(* IEC 61131-3 sources: volt/packages/volt-lsp-iec/test-corpus/bakon-nano/Device/Plc Logic/Application/Library Manager/L_TS2P_TechModulesSynchronizingCamming (part 2) *)

(* ---- L_TS2P_CALCULATETARGETPOS.pou ---- *)
FUNCTION_BLOCK L_TS2P_CALCULATETARGETPOS
VAR_INPUT
	XRESET : BOOL;
	XENABLE : BOOL;
	XEXECUTENEXTCUT : BOOL;
	XEXECUTEFIRSTCUT : BOOL;
	XSETCUTTINGLENGTHINSTANT : BOOL;
	XTPNOTVALID : BOOL;
	XEXECUTEGAP : BOOL;
	XRESUMETARGETPOS : BOOL;
	XSTARTFLYINGSAW : BOOL;
	ETMSTATE : L_TB2P_States;
	XSYNCININSTANT : BOOL;
	XSETMATERIALCOUNTER : BOOL;
	LRMATERIALCOUNTER : LREAL;
	LRDELTAMATERIALPOS : LREAL;
	LRSLAVEPOS : LREAL;
	LRCUTTINGLENGTH : LREAL;
	LRMARKSENSORPOS : LREAL;
	LRGAP : LREAL;
	LRMARKPOSITION : LREAL;
	XLOADTOTALCUTTINGLENGTH : BOOL;
	LRLOADTOTALCUTTINGLENGTH : LREAL;
	XLOADTARGETPOS : BOOL;
	LRLOADTARGETPOS : LREAL;
	EMODE : L_TS2P_FlyingSawMode;
	LRVELINMASTER : LREAL;
	LRACCDIST : LREAL;
	LRACCTIME : LREAL;
	LRTASKCYCLETIME : LREAL;
	XEMPTYSTACK : BOOL;
	XSYNCHRONIZED : BOOL;
	XINPOSITION : BOOL;
END_VAR
VAR_OUTPUT
	XEXECUTEGAPOUT : BOOL;
	LRTARGETPOS : LREAL;
	LRTARGETPOS_OUT : LREAL;
	LRTOTALPRODUCTLENGTH : LREAL;
	XCUTTINGLENGTHVALID : BOOL;
	LRACTIVECUTTINGLENGTH : LREAL;
END_VAR
VAR
	LROFFSET_INT : LREAL;
	XGAPREQUESTED : BOOL;
	LRDELTAMATERIALPOS_INT : LREAL;
	LRTOLERANCE : LREAL;
	LROFFSETOUT_INT : LREAL;
	LRGAPTOTAL_INT : LREAL;
	XSYNCININSTANT_LOCK : BOOL;
	XENABLE_OLD : BOOL;
	XSYNCININSTANT_OLD : BOOL;
	LRMATERIALCOUNTER_OLD : LREAL;
	XEXECUTENEXTCUT_OLD : BOOL;
	XEXECUTEGAP_OLD : BOOL;
	XEXECUTEFIRSTCUT_OLD : BOOL;
	EMODE_OLD : WORD;
	ETMSTATE_OLD : L_TB2P_States;
	XTPNOTVALID_OLD : BOOL;
	XSETCUTTINGLENGTHINSTANT_OLD : BOOL;
	XSETMATERIALCOUNTER_OLD : BOOL;
	LRMARKPOSITION_OLD : LREAL;
END_VAR
END_FUNCTION_BLOCK

(* ---- L_TS2P_CALCULATETPCOMPENSATIONFACTOR.pou ---- *)
FUNCTION_BLOCK L_TS2P_CALCULATETPCOMPENSATIONFACTOR
VAR_OUTPUT
	LRFACTOR : LREAL;
	LRCOMPENSATIONCYCLES : LREAL;
END_VAR
VAR_IN_OUT
	TPAXIS : AXIS_REF;
END_VAR
VAR
	LRSETPOSARRAY : ARRAY [0..15] OF LREAL;
	BYCOUNTER : BYTE;
	LRTEMP : LREAL;
	LRPOSDIFF : LREAL;
	LRSETACTDIFF : LREAL;
	XERRORINVALIDAXIS : BOOL;
	LRSETPOS : LREAL;
	LRACTPOS : LREAL;
	LRCYCLELENGTH : LREAL;
	LRADDITIONALCORRECTION : LREAL;
	LRTEMP2 : LREAL;
	XINCREMENTCYCLES : BOOL;
END_VAR
END_FUNCTION_BLOCK

METHOD SEARCHARRAY
END_METHOD

(* ---- L_TS2P_CALCULATETPONMATERIALPOS.pou ---- *)
FUNCTION_BLOCK L_TS2P_CALCULATETPONMATERIALPOS
VAR_INPUT
	XENABLE : BOOL;
	BYTASKCYCLEDELAY : BYTE := 4;
	XMARKRECEIVE : BOOL;
	LRMARKSENSORPOS : LREAL;
	LRACTMARKPOSIN : LREAL;
	LRCYCPOSTPAXIS : LREAL;
	LRCYCVELTPAXIS : LREAL;
	LRCYCLELENGTHTPAXIS : LREAL;
	LRCYCLELENGTHTARGETAXIS : LREAL;
	LRTASKCYCLETIME : LREAL;
	XRESETMARKSTACK : BOOL;
	LRMATERIALCOUNTER : LREAL;
	LRUPPERLIMITWORKINGRANGE : LREAL;
	LRLOWERLIMITWORKINGRANGE : LREAL;
	LRFACTOR : LREAL;
	LRCOMPVELFACTOR : LREAL;
	XSCIPTONEXTPOSOUT : BOOL;
	XSYNCININSTANT : BOOL;
	XEXECUTEFIRSTCUT : BOOL;
END_VAR
VAR_OUTPUT
	LRTPPOSOUT : LREAL;
	XEXECUTEFIRSTCUT_OLD : BOOL;
	LRTPACTTIMESTAMP : LREAL;
	XFULL : BOOL;
	WMARKPOSITIONVALID : WORD;
	WININDEX : WORD;
	ALRMARKPOSITIONARRAY : ARRAY [0..15] OF LREAL := [0, 0, 0, 0, 0, 0, 0, 0, 0, 0, 0, 0, 0, 0, 0, 0];
	ALRTIMESTAMPARRAY : ARRAY [0..15] OF LREAL;
	XEMPTY : BOOL := TRUE;
	WOUTINDEX : WORD;
	BYREMAINMARKSTACK : BYTE := 15;
	XTPRECEIVED : BOOL;
	XMARKRECEIVED : BOOL;
	XTPPOSVALID : BOOL;
	BYCOUNTEROUT : BYTE;
	XERROR : BOOL;
END_VAR
VAR
	R_TRIG1 : R_TRIG;
	LRTIMESTAMP : LREAL;
	BYTPIDLEINDEX : BYTE;
	BYTPACTINDEX : BYTE;
	ALRPOSITION : ARRAY [0..15] OF LREAL;
	BYTPPREVINDEX : BYTE;
	BYTMP : BYTE;
	XSKIPTONEXTPOS : BOOL;
	WTESTCOUNTER : WORD;
	XTEST : BOOL;
	XWAIT : BOOL;
	WCOUNTINVALIDTIMESTAMP : WORD;
	LRDISTINACTMASTER : LREAL;
	BYTEST : BYTE;
	LRMARKPOSITIONDIFF : LREAL;
	LRMARKPOSITIONDIFF2 : LREAL;
	LRPOSFIFOX : ARRAY [1..20] OF LREAL := [10(0)];
	LRPOSFIFOREG : ARRAY [1..20] OF LREAL := [10(0)];
	BYCOUNTER : BYTE := 1;
	LRSTACKDIFFERENCE : LREAL;
	LRTPDELTAINMS : LREAL;
	LRDELTAPCT : LREAL;
	LRTEMP : LREAL;
	IDIRECTION : INT;
	LRACTMARKPOSIN_OLD : LREAL;
	R_TRIG2 : R_TRIG;
	DWSTATE : DWORD;
	WSTOREDPOSVALUES : WORD;
	LRACTMARKPOSIN_INT : LREAL;
	XSYNCININSTANT_OLD : BOOL;
	XWAIT_OLD : BOOL;
	XRESETMARKSTACK_OLD : BOOL;
	BYCNT : BYTE;
	BYSTEPPER : BYTE;
END_VAR
END_FUNCTION_BLOCK

METHOD SEARCHINSTACKNEGATIVE
END_METHOD

METHOD SEARCHINSTACKPOSITIVE
END_METHOD

(* ---- L_TS2P_CAMCREATOR.pou ---- *)
FUNCTION_BLOCK L_TS2P_CAMCREATOR
VAR_INPUT
	XENABLEINTERNALCAMTABLE : BOOL;
	XEXECUTE : BOOL;
	PCAMPOINTS : POINTER TO L_MC2P_CamDataXYVA;
	INUMOFPOINTS : INT;
	LRMASTERMAXVEL : LREAL;
	LRMASTERMAXACC : LREAL;
	LRMASTERSCALING : LREAL := 1;
	LRSLAVESCALING : LREAL := 1;
END_VAR
VAR_OUTPUT
	XINTERNALCAMTABLELACTIVE : BOOL;
	XERROR : BOOL;
	EERRORID : L_IE1P_Error;
	XBUSY : BOOL;
	XDONE : BOOL;
	CAMTABLEOUT : MC_CAM_REF;
	LRSLAVEMAXPOS : LREAL;
	LRSLAVEMINPOS : LREAL;
	LRSLAVEMAXVEL : LREAL;
	LRSLAVEMINVEL : LREAL;
	LRSLAVEMAXACC : LREAL;
	LRSLAVEMINACC : LREAL;
END_VAR
VAR_IN_OUT
	SLAVE : AXIS_REF;
END_VAR
VAR
	EFMSTATE : L_MB1P_States := L_MB1P_States.INIT;
	SMC_CAMBOUNDS1 : L_MC2P_BoundsCam;
	SMC_CAMBOUNDSINIT : L_MC2P_BoundsCam;
	CAMREF : L_MC2P_CamRefFromStruct;
	PCAMPOINTS_INT : POINTER TO L_MC2P_CamDataXYVA;
	INUMOFPOINTS_INT : INT;
	XINTERNALCONTROL : BOOL;
	XEXECUTE_OLD : BOOL;
	ASCCAMPOINTS : ARRAY [0..30] OF L_MC2P_CamDataXYVA;
	XINVALIDCAMTABLE : BOOL;
	XVISUACTIVE : BOOL := TRUE;
	DIFRAME : DINT;
	DIFRAME_OLD : DINT;
	ARVISPOINTLINES : ARRAY [1..10] OF L_MC2P_CamDataXYVA;
	IVISUTABLESETPOS : INT := 0;
	IVISUTABLESETPOS_OLD : INT := 0;
	IVISUTABLEMAXPOS : INT := 30;
	IVISSHOWLINESNO : INT;
	XVISPOINTMIN : BOOL;
	XVISPOINTMAX : BOOL;
	XVISUSETPOSUP : BOOL;
	XVISUSETPOSDOWN : BOOL;
	XVISUSETPOSUP_OLD : BOOL;
	XVISUSETPOSDOWN_OLD : BOOL;
	XSCROLBUTTENACTIVE : BOOL;
	TSETTIME : TIME := TIME#400ms;
	TON_SCROLBUTTEN : TON;
END_VAR
END_FUNCTION_BLOCK

METHOD CALL_CAMBOUNDS
VAR_IN_OUT
	SLAVE : AXIS_REF;
END_VAR
END_METHOD

METHOD CALL_CAMREF
END_METHOD

METHOD CALL_CAMTABLEEQUIDISTANT
END_METHOD

METHOD CALL_CAMTABLENONEQUIDISTANT
END_METHOD

METHOD CALL_CAMTABLEPOLYNOMIAL
END_METHOD

METHOD CALL_ERRORHANDLER
END_METHOD

METHOD CALL_FBMETHODS
VAR_IN_OUT
	SLAVE : AXIS_REF;
END_VAR
END_METHOD

METHOD CALL_INTERNALCTRL
END_METHOD

METHOD CALL_OUTPUT
END_METHOD

METHOD CALL_RESETCOMMANDS
VAR_IN_OUT
	SLAVE : AXIS_REF;
END_VAR
END_METHOD

METHOD CALL_RESETOUTPUT
END_METHOD

METHOD CALL_STATEMACHINE
END_METHOD

METHOD CALL_VIS_TON_SCROLBUTTEN
END_METHOD

METHOD CALL_VISUTABCTRL
END_METHOD

METHOD CALL_VISUUPDATETAB
END_METHOD

METHOD DISABALE_VISU
END_METHOD

METHOD ENABLE_VISU
END_METHOD

METHOD CALL_S000_CYCLIC
END_METHOD

METHOD CALL_S001_INIT
END_METHOD

METHOD CALL_S002_READY
END_METHOD

(* ---- L_TS2P_CAMTABLEINFO.pou ---- *)
FUNCTION_BLOCK L_TS2P_CAMTABLEINFO
VAR_INPUT
	XENABLE : BOOL;
	CAMTABLE : MC_CAM_REF;
	LRMASTERMAXVEL : LREAL := 100;
	LRMASTERMAXACC : LREAL := 1000;
	LRMASTERSCALING : LREAL := 1;
	LRSLAVESCALING : LREAL := 1;
END_VAR
VAR_OUTPUT
	XBUSY : BOOL;
	XDONE : BOOL;
	XCAMTABLEVALID : BOOL;
	LRMASTERSTARTPOS : LREAL;
	LRMASTERENDPOS : LREAL;
	LRSLAVESTARTPOS : LREAL;
	LRSLAVEENDPOS : LREAL;
	LRSLAVEMAXPOS : LREAL;
	LRSLAVEMINPOS : LREAL;
	LRSLAVEMAXVEL : LREAL;
	LRSLAVEMINVEL : LREAL;
	LRSLAVEMAXACC : LREAL;
	LRSLAVEMINACC : LREAL;
END_VAR
VAR_IN_OUT
	SLAVEAXIS : AXIS_REF;
END_VAR
VAR
	ESTATE : L_MB1P_States := L_MB1P_States.INIT;
	CAMTABLE_INT : MC_CAM_REF;
	PCAMDATA_INT : POINTER TO L_MC2P_CamData;
	LRMASTERMAXVEL_INT : LREAL := 0;
	LRMASTERMAXACC_INT : LREAL := 0;
	LRMASTERSCALING_INT : LREAL := 0;
	LRSLAVESCALING_INT : LREAL := 0;
	XENABLE_OLD : BOOL;
	SMC_CAMBOUNDS1 : L_MC2P_BoundsCam;
	XCALCNEWVALUES : BOOL;
END_VAR
END_FUNCTION_BLOCK

METHOD CALC_STARTENDVALUES
END_METHOD

METHOD CALL_CAMBOUNDS
END_METHOD

METHOD CALL_FBMETHODS
END_METHOD

METHOD CALL_OUTPUT
END_METHOD

METHOD CALL_RESETCOMMANDS
END_METHOD

METHOD CALL_RESETOUTPUT
END_METHOD

METHOD CALL_STATEMACHINE
END_METHOD

METHOD GET_XCALCNEWVALUES : BOOL
END_METHOD

METHOD GET_XCRITICALCYCLE : BOOL
END_METHOD

(* ---- L_TS2P_CONDITIONLIMITERSYNCIN.pou ---- *)
FUNCTION_BLOCK L_TS2P_CONDITIONLIMITERSYNCIN EXTENDS L_UBUP_ConditionBase
VAR_INPUT
	ESYNCDIRECTION : L_TS2P_SyncDirection;
	DWLIMITERCONTROL : DWORD;
END_VAR
VAR_OUTPUT
	XDIRECTIONDISABLED : BOOL;
	XINVALIDINPUT : BOOL;
END_VAR
VAR_IN_OUT
	AXIS : AXIS_REF;
END_VAR
END_FUNCTION_BLOCK

METHOD VERIFY : BOOL
VAR_OUTPUT
	XCONDITIONERROR : BOOL;
	EERRORIDPROPOSED : L_IE1P.L_IE1P_Error;
END_VAR
END_METHOD

(* ---- L_TS2P_CONDITIONLOCKTOCAM.pou ---- *)
FUNCTION_BLOCK L_TS2P_CONDITIONLOCKTOCAM EXTENDS L_UBUP_ConditionBase
VAR_IN_OUT
	SCPAR : L_TS2P_scPar_TM_FlexCam;
END_VAR
END_FUNCTION_BLOCK

METHOD VERIFY : BOOL
VAR_OUTPUT
	XCONDITIONERROR : BOOL;
	EERRORIDPROPOSED : L_IE1P.L_IE1P_Error;
END_VAR
END_METHOD

(* ---- L_TS2P_CONDITIONSYNCPARAMETER.pou ---- *)
FUNCTION_BLOCK L_TS2P_CONDITIONSYNCPARAMETER EXTENDS L_UBUP_ConditionBase
VAR_IN_OUT
	SCPAR : L_TS2P_scPar_TM_SyncPosBase;
END_VAR
END_FUNCTION_BLOCK

METHOD VERIFY : BOOL
VAR_OUTPUT
	XCONDITIONERROR : BOOL;
	EERRORIDPROPOSED : L_IE1P.L_IE1P_Error;
END_VAR
END_METHOD

(* ---- L_TS2P_CONDITIONVALIDCAMTABLE.pou ---- *)
FUNCTION_BLOCK L_TS2P_CONDITIONVALIDCAMTABLE EXTENDS L_UBUP_ConditionBase
VAR_INPUT
	WSETCAMTABLE : WORD;
	CAMTABLE1 : MC_CAM_REF;
	CAMTABLE2 : MC_CAM_REF;
	CAMTABLE3 : MC_CAM_REF;
	CAMTABLE4 : MC_CAM_REF;
END_VAR
END_FUNCTION_BLOCK

METHOD VERIFY : BOOL
VAR_OUTPUT
	XCONDITIONERROR : BOOL;
	EERRORIDPROPOSED : L_IE1P.L_IE1P_Error;
END_VAR
END_METHOD

(* ---- L_TS2P_CROSSCUTTERSTATE.pou ---- *)
FUNCTION_BLOCK L_TS2P_CROSSCUTTERSTATE EXTENDS L_TB2P_TechModuleBase
VAR_INPUT
	XENABLE : BOOL;
	XENABLEOPERATION : BOOL;
	XRESETERROR : BOOL;
	XQSPAPPLICATION : BOOL;
	XABORT : BOOL;
	XJOGPOS : BOOL;
	XJOGNEG : BOOL;
	XHOMEEXECUTE : BOOL;
	LROVERRIDE : LREAL := 1;
	SCCTRLBASICMOTION : L_TB2P_scCtrlBasicMotion;
	SCPAR : L_TS2P_scPar_CrossCutterState;
	SCACCESSPOINTS : L_TS2P_scAP_CrossCutterState;
	MASTERVALUES : L_MC1P_IAXIS_REF_MASTERVALUES;
	XEXECUTEMOVETOPARKPOS : BOOL;
	XSYNCIN : BOOL;
	XHOLDINPARKPOS : BOOL;
	LRPRODUCTLENGTH : LREAL;
	LROVERSPEED : LREAL;
	LRSETOFFSETPOSX : LREAL;
	XTRIMPOS : BOOL;
	XTRIMNEG : BOOL;
	XTRIMRESET : BOOL;
	SCTPRECDATA_MARKSENSOR : L_MC1P_TpReceiveData;
	SCTPRECDATA_TOOLSENSOR : L_MC1P_TpReceiveData;
	XTEACHMARKWINDOW : BOOL;
	XTEACHMARKWINDOWTOOL : BOOL;
	XGEARFACTORCORR : BOOL;
	XGEARFACTORCORRHOLD : BOOL;
END_VAR
VAR_OUTPUT
	XREADYFOROPERATION : BOOL;
	XOPERATIONENABLED : BOOL;
	XREADYFORMOTION : BOOL;
	XERROR : BOOL;
	XWARNING : BOOL;
	EERRORID : L_IE1P_Error;
	XSTOACTIVE : BOOL;
	XQSPACTIVE : BOOL;
	XABORTBUSY : BOOL;
	XABORTDONE : BOOL;
	XJOGGINGBUSY : BOOL;
	XHOMINGBUSY : BOOL;
	XHOMINGDONE : BOOL;
	XISHOMED : BOOL;
	ETMSTATE : L_TB2P_States;
	SCSTATUSBASICMOTION : L_TB2P_scStatusBasicMotion;
	LRACTVEL : LREAL;
	LRSETVELOUT : LREAL;
	LRACTPOS : LREAL;
	LRSETPOSOUT : LREAL;
	LRACTFOLLOWINGERROR : LREAL;
	SCSIGNALFLOW : L_TS2P_scSF_CrossCutterState;
	XSYNCHRONISED : BOOL;
	XACCDECSYNC : BOOL;
	XOFFSETTRIMACTIVE : BOOL;
	XINPARKPOS : BOOL;
	XHOLDINPARKPOSACTIVE : BOOL;
	XCUTDONE : BOOL;
	XCUTTINGACTIVE : BOOL;
	LRACTCUTLENGTH : LREAL;
	LROFFSETTOTAL : LREAL;
	XTRQCTRLACTIVE : BOOL;
	LRSETMARKCORROUT : LREAL;
	XMARKWINDOWTEACHED : BOOL;
	LRGEARFACTORCORR : LREAL;
	LRSETTOOLCORROUT : LREAL;
	XMARKWINDOWTEACHEDTOOL : BOOL;
END_VAR
VAR_IN_OUT
	AXIS : AXIS_REF;
END_VAR
VAR
	TM_INT : L_TS2P_TM_CrossCutterState := STRUCT(ModuleHandler := ModuleHandler);
	SCPAR_INT : L_TS2P_scPar_CrossCutterState;
	_UICALLMFUNIDXINPUT : UINT := 1;
	_UICALLMFUNIDXOUTPUT : UINT := 1;
	_MCCALL : L_UM1P_MCCall;
	_ASCINPUT : ARRAY [1.._MCCall.c_BufferDepthInput] OF L_TS2P_CrossCutterStateIn;
	_ASCOUTPUT : ARRAY [1.._MCCall.c_BufferDepthOutput] OF L_TS2P_CrossCutterStateOut;
	_ASCPARCORE : ARRAY [1.._MCCall.c_BufferDepthInput] OF L_TS2P_scPar_CrossCutterState;
	_ASCACCESSPOINTSCORE : ARRAY [1.._MCCall.c_BufferDepthInput] OF L_TS2P_scAP_CrossCutterState;
	_ASCSIGNALFLOWCORE : ARRAY [1.._MCCall.c_BufferDepthOutput] OF L_TS2P_scSF_CrossCutterState;
	_SCINPUTVISU : L_TS2P_CrossCutterStateIn;
	_PSCINPUTVISU : POINTER TO L_TS2P_CrossCutterStateIn := ADR(_scInputVisu);
	_PSCOUTPUTVISU : POINTER TO L_TS2P_CrossCutterStateOut := ADR(_ascOutput[1]);
	_PSCPARVISU : POINTER TO L_TS2P_scPar_CrossCutterState := ADR(scPar_int);
	ITFITECHMODULEINTERNAL : L_TB2P_ITechModuleInternal;
	LRJERKDEC : LREAL;
	LRJOGGINGJERKDEC : LREAL;
	REMAININGTIMEOFPROFILE : LREAL;
	REMAININGTIMEOFPROFILEAVAILABLE : BOOL;
END_VAR
END_FUNCTION_BLOCK

METHOD GET_PAP : POINTER TO L_TB2P_scAP_TM_MotionControl
END_METHOD

METHOD GET_PPAR : POINTER TO L_TB2P_scPar_TM_MotionControl
END_METHOD

METHOD GET_PSF : POINTER TO L_TB2P_scSF_TM_MotionControl
END_METHOD

METHOD CALLFUNCTION
VAR_INPUT
	UIINPUTDATAIDX : UINT;
	UIOUTPUTDATAIDX : UINT;
END_VAR
END_METHOD

METHOD COPYINPUTS : BOOL
VAR_INPUT
	IDX : WORD;
END_VAR
END_METHOD

METHOD COPYOUTPUTS : BOOL
VAR_INPUT
	IDX : WORD;
END_VAR
END_METHOD

METHOD FUNCTIONWASCALLEDTWICE : BOOL
VAR_INPUT
	IDX : WORD;
END_VAR
END_METHOD

METHOD HANDLESTANDARDCALL : BOOL
END_METHOD

METHOD SYNCOUTPUTS
VAR_INPUT
	UICOPYOUTPUTFROMIDX : UINT;
	UICOPYOUTPUTTOIDX : UINT;
END_VAR
END_METHOD

METHOD CALL_INTERNALCTRL
END_METHOD

(* ---- L_TS2P_DISTCORRECTIONWINDOW.pou ---- *)
FUNCTION_BLOCK L_TS2P_DISTCORRECTIONWINDOW
VAR_INPUT
	XENABLE : BOOL;
	XENABLEPOSITION : BOOL;
	LRCYCSETPOSMASTER : LREAL;
	LRCYCLELENGTHMASTER : LREAL;
	LRCYCSETVEL : LREAL;
	XLOADSTARTPOS : BOOL;
	LRSTARTPOS : LREAL;
	XTPRECEIVEDIN : BOOL;
	LRSETCORRECTION : LREAL;
	XCORRWINDOWINXUNITS : BOOL;
	LRSETUPPERWINDOW : LREAL;
	LRSETLOWERWINDOW : LREAL;
	LRCYCPOSFEEDBACK : LREAL;
	DNSETNUMERATORAXISY : DWORD := 1;
	DNSETDENOMINATORAXISY : DWORD := 1;
	LRSETCYCLELENGTHX : LREAL;
	LRSETCYCLELENGTHY : LREAL;
END_VAR
VAR_OUTPUT
	XBUSY : BOOL;
	XCORRECTIONBUSY : BOOL;
	LRSETPOSOUT : LREAL;
	LRSETINTEGRATEDPOSITION : LREAL;
	LRSETPOSCORROUT : LREAL;
	LRSETPOSCORRRESIDUALOUT : LREAL;
	LRDELTAPOSCORROUT : LREAL;
	XCORRNEXTCYCLE : BOOL;
	XERROR : BOOL;
	EERRORID : L_IE1P_Error;
END_VAR
VAR
	LRDELTAPOSTOTAL : LREAL;
	LRMASTERDISTANCE : LREAL;
	LRPOSITIONSET : LREAL;
	LRPOSITIONNORMED : LREAL;
	LRPOSITIONOUTNORMED : LREAL;
	LRDELTAPOSCORRECTION : LREAL;
	LRPOSITIONSETOLD : LREAL;
	LRPOSITIONSETAXISOUT : LREAL;
	BYSTEPPER : BYTE;
	LRCORRECTIONDISTANCELOCAL : LREAL;
	LRCORRECTIONLOCAL : LREAL;
	L_DIFFERENTIATE : L_MC2P_Differentiate;
	INTEGRATOR : L_MC1P_IntegrateAxis;
	LRDELTAPOSOUT : LREAL;
	XEXECUTECORRECTIONINTERN : BOOL;
	XPOSITIVEDIRECTION : BOOL := FALSE;
	LRCORRECTIONDISTANCE : LREAL;
	LRUPPERWINDOWINTERNAL : LREAL;
	LRLOWERWINDOWINTERNAL : LREAL;
	LRTASKCYCLE : LREAL;
	XCORRECTIONACTIVE : BOOL;
	LRCORRECTIONLOCAL1 : LREAL;
	XTPRECEIVEDOLD : BOOL;
	LRINTEGRATORSPEED : LREAL;
	XWINDOWINCYCLE : BOOL;
	LRDELTAWINDOW : LREAL;
	LRCYCPOSINTOOLINTERNAL : LREAL;
	LRUPPERWINDOWINTERNALDELTA : LREAL;
	LRLOWERWINDOWINTERNALDELTA : LREAL;
	XINIT : BOOL := TRUE;
	XINITOUTOFCORRWINDOW : BOOL := TRUE;
	LRLOWERWINDOWINTERNALOLD : LREAL;
	LRUPPERWINDOWINTERNALOLD : LREAL;
	LRCYCPOSFEEDBACKINT : LREAL;
	XCORRECTIONBUSYOLD : BOOL;
	LRSETPOSCORROUTOLD : LREAL;
	LRCYCPOSINTOOLINTERNAL_CASE : LREAL;
	XWINDOWCHANGEDFLAG : BOOL := FALSE;
	LRCYCLELENGTH_INT : LREAL;
	LROFFSET_INT : LREAL;
	LRCYCPOSINTOOLINTERNAL_0LD : LREAL;
	LRPOSITIONNORMED_OLD : LREAL;
	LRPOSITIONNORMED_DIF : LREAL;
	XPOSCORR : BOOL;
	XTPSTORED_INT : BOOL;
	LRSETCORRECTIONSTORED_INT : LREAL;
	XINCORRWINDOW : BOOL;
	XINCORRWINDOWOLD : BOOL;
	LRSETPOSOUTCOMP : LREAL;
	LRCYCPOSINTOOLINTERNALOLD : LREAL;
	LRDELTAPOSOUTINTERNAL : LREAL;
	BYSTEPPEROLD : BYTE := 0;
	LRCYCSETPOSOLD : LREAL;
	LRCORRECTIONINYUNITS : LREAL;
	LRCORRECTIONDISTANCETEMP : LREAL;
END_VAR
END_FUNCTION_BLOCK

METHOD CALL_INIT
END_METHOD

(* ---- L_TS2P_ELECTRONICGEARBOXBASE.pou ---- *)
FUNCTION_BLOCK L_TS2P_ELECTRONICGEARBOXBASE EXTENDS L_TB2P_TechModuleBase
VAR_INPUT
	XENABLE : BOOL;
	XENABLEOPERATION : BOOL;
	XRESETERROR : BOOL;
	XQSPAPPLICATION : BOOL;
	XABORT : BOOL;
	XJOGPOS : BOOL;
	XJOGNEG : BOOL;
	XHOMEEXECUTE : BOOL;
	LROVERRIDE : LREAL := 1;
	SCCTRLBASICMOTION : L_TB2P_scCtrlBasicMotion;
	SCPAR : L_TS2P_scPar_ElectronicGearboxBase;
	SCACCESSPOINTS : L_TS2P_scAP_ElectronicGearboxBase;
	MASTERVALUES : L_MC1P_IAXIS_REF_MASTERVALUES;
	XSYNCIN : BOOL;
	LRSETBASEVEL : LREAL;
	LRSETOFFSETPOS : LREAL;
	LRSETOFFSETVEL : LREAL;
	XTRIMPOS : BOOL;
	XTRIMNEG : BOOL;
	XTRIMRESET : BOOL;
	XINVERTGEARFACTOR : BOOL;
END_VAR
VAR_OUTPUT
	XREADYFOROPERATION : BOOL;
	XOPERATIONENABLED : BOOL;
	XREADYFORMOTION : BOOL;
	XERROR : BOOL;
	XWARNING : BOOL;
	EERRORID : L_IE1P_Error;
	XSTOACTIVE : BOOL;
	XQSPACTIVE : BOOL;
	XABORTBUSY : BOOL;
	XABORTDONE : BOOL;
	XJOGGINGBUSY : BOOL;
	XHOMINGBUSY : BOOL;
	XHOMINGDONE : BOOL;
	XISHOMED : BOOL;
	ETMSTATE : L_TB2P_States := L_TB2P_States.DISABLED;
	SCSTATUSBASICMOTION : L_TB2P_scStatusBasicMotion;
	LRACTVEL : LREAL;
	LRSETVELOUT : LREAL;
	LRACTPOS : LREAL;
	LRSETPOSOUT : LREAL;
	LRACTFOLLOWINGERROR : LREAL;
	SCSIGNALFLOW : L_TS2P_scSF_ElectronicGearboxBase;
	XSYNCHRONISED : BOOL;
	XACCDECSYNC : BOOL;
	XOFFSETTRIMACTIVE : BOOL;
	XBASEVELOCITYACTIVE : BOOL;
	LROFFSETTOTALVEL : LREAL;
END_VAR
VAR_IN_OUT
	AXIS : AXIS_REF;
END_VAR
VAR
	TM_INT : L_TS2P_TM_ElectronicGearboxBase := STRUCT(ModuleHandler := ModuleHandler);
	SCPAR_INT : L_TS2P_scPar_ElectronicGearboxBase;
	_UICALLMFUNIDXINPUT : UINT := 1;
	_UICALLMFUNIDXOUTPUT : UINT := 1;
	_MCCALL : L_UM1P_MCCall;
	_ASCINPUT : ARRAY [1.._MCCall.c_BufferDepthInput] OF L_TS2P_ElectronicGearboxBaseIn;
	_ASCOUTPUT : ARRAY [1.._MCCall.c_BufferDepthOutput] OF L_TS2P_ElectronicGearboxBaseOut;
	_ASCPARCORE : ARRAY [1.._MCCall.c_BufferDepthInput] OF L_TS2P_scPar_ElectronicGearboxBase;
	_ASCACCESSPOINTSCORE : ARRAY [1.._MCCall.c_BufferDepthInput] OF L_TS2P_scAP_ElectronicGearboxBase;
	_ASCSIGNALFLOWCORE : ARRAY [1.._MCCall.c_BufferDepthOutput] OF L_TS2P_scSF_ElectronicGearboxBase;
	_SCINPUTVISU : L_TS2P_ElectronicGearboxBaseIn;
	_PSCINPUTVISU : POINTER TO L_TS2P_ElectronicGearboxBaseIn := ADR(_scInputVisu);
	_PSCOUTPUTVISU : POINTER TO L_TS2P_ElectronicGearboxBaseOut := ADR(_ascOutput[1]);
	_PSCPARVISU : POINTER TO L_TS2P_scPar_ElectronicGearboxBase := ADR(scPar_int);
	ITFITECHMODULEINTERNAL : L_TB2P_ITechModuleInternal;
	LRJERKDEC : LREAL;
	LRJOGGINGJERKDEC : LREAL;
	REMAININGTIMEOFPROFILE : LREAL;
	REMAININGTIMEOFPROFILEAVAILABLE : BOOL;
END_VAR
END_FUNCTION_BLOCK

METHOD GET_PAP : POINTER TO L_TB2P_scAP_TM_MotionControl
END_METHOD

METHOD GET_PPAR : POINTER TO L_TB2P_scPar_TM_MotionControl
END_METHOD

METHOD GET_PSF : POINTER TO L_TB2P_scSF_TM_MotionControl
END_METHOD

METHOD CALLFUNCTION
VAR_INPUT
	UIINPUTDATAIDX : UINT;
	UIOUTPUTDATAIDX : UINT;
END_VAR
END_METHOD

METHOD COPYINPUTS : BOOL
VAR_INPUT
	IDX : WORD;
END_VAR
END_METHOD

METHOD COPYOUTPUTS : BOOL
VAR_INPUT
	IDX : WORD;
END_VAR
END_METHOD

METHOD FUNCTIONWASCALLEDTWICE : BOOL
VAR_INPUT
	IDX : WORD;
END_VAR
END_METHOD

METHOD HANDLESTANDARDCALL : BOOL
END_METHOD

METHOD SYNCOUTPUTS
VAR_INPUT
	UICOPYOUTPUTFROMIDX : UINT;
	UICOPYOUTPUTTOIDX : UINT;
END_VAR
END_METHOD

METHOD CALL_INTERNALCTRL
END_METHOD

(* ---- L_TS2P_FLEXCAMHIGH.pou ---- *)
FUNCTION_BLOCK L_TS2P_FLEXCAMHIGH EXTENDS L_TB2P_TechModuleBase
VAR_INPUT
	XUSEORIGINAL : BOOL;
	XENABLE : BOOL;
	XENABLEOPERATION : BOOL;
	XRESETERROR : BOOL;
	XQSPAPPLICATION : BOOL;
	XABORT : BOOL;
	XJOGPOS : BOOL;
	XJOGNEG : BOOL;
	XHOMEEXECUTE : BOOL;
	LROVERRIDE : LREAL := 1;
	SCCTRLBASICMOTION : L_TB2P_scCtrlBasicMotion;
	SCPAR : L_TS2P_scPar_FlexCamHigh;
	SCACCESSPOINTS : L_TS2P_scAP_FlexCamHigh;
	MASTERVALUES : L_MC1P_IAXIS_REF_MASTERVALUES;
	XCLUTCHCLOSE : BOOL;
	XLOADCLUTCHPOS : BOOL;
	LRLOADCLUTCHPOS : LREAL;
	XFINDCLUTCHXPOS : BOOL;
	XSYNCIN : BOOL;
	XSYNCPOSRESTORE : BOOL;
	XCAMCHANGEINSTANT : BOOL;
	LRSETOFFSETPOSX : LREAL;
	LRSETOFFSETPOSY : LREAL;
	LRSETSCALINGX : LREAL := 1;
	LRSETSCALINGY : LREAL := 1;
	CAMTABLE1 : MC_CAM_REF;
	CAMTABLE2 : MC_CAM_REF;
	CAMTABLE3 : MC_CAM_REF;
	CAMTABLE4 : MC_CAM_REF;
	WSETCAMTABLE : WORD := 1;
	XCAMSEQUENCER : BOOL;
END_VAR
VAR_OUTPUT
	XREADYFOROPERATION : BOOL;
	XOPERATIONENABLED : BOOL;
	XREADYFORMOTION : BOOL;
	XERROR : BOOL;
	XWARNING : BOOL;
	EERRORID : L_IE1P_Error;
	XSTOACTIVE : BOOL;
	XQSPACTIVE : BOOL;
	XABORTBUSY : BOOL;
	XABORTDONE : BOOL;
	XJOGGINGBUSY : BOOL;
	XHOMINGBUSY : BOOL;
	XHOMINGDONE : BOOL;
	XISHOMED : BOOL;
	ETMSTATE : L_TB2P_States;
	SCSTATUSBASICMOTION : L_TB2P_scStatusBasicMotion;
	LRACTVEL : LREAL;
	LRSETVELOUT : LREAL;
	LRACTPOS : LREAL;
	LRSETPOSOUT : LREAL;
	LRACTFOLLOWINGERROR : LREAL;
	SCSIGNALFLOW : L_TS2P_scSF_FlexCamHigh;
	XCLUTCHACTIVE : BOOL;
	XCLUTCHCLOSED : BOOL;
	XACCDECSYNC : BOOL;
	XSYNCHRONISED : BOOL;
	XMOVETOPARKPOSACTIVE : BOOL;
	XINPARKPOS : BOOL;
	XENDOFPROFILE : BOOL;
	LROFFSETPOSX : LREAL;
	LROFFSETPOSY : LREAL;
	LROFFSETSYNCPOS : LREAL;
	WACTIVECAMTABLE : WORD;
	XCAMSEQUENCERACTIVE : BOOL;
END_VAR
VAR_IN_OUT
	AXIS : AXIS_REF;
END_VAR
VAR
	XINTERNALCONTROLACTIVE_OLD : BOOL;
	ITFCONNECTORFLEXCAM : L_TS2P_IConnectorFlexCam;
	TM_INT : L_TS2P_TM_FlexCam;
	SCPAR_INT : L_TS2P_scPar_FlexCamHigh;
	SCDATA_INT : L_TS2P_scData_TM_FlexCam;
	SCDATASP_INT : L_TS2P_scData_TM_FlexCam;
	XUSEORIGINAL_OLD : BOOL;
	_UICALLMFUNIDXINPUT : UINT := 1;
	_UICALLMFUNIDXOUTPUT : UINT := 1;
	_MCCALL : L_UM1P_MCCall;
	_ASCINPUT : ARRAY [1.._MCCall.c_BufferDepthInput] OF L_TS2P_FlexCamHighIn;
	_ASCOUTPUT : ARRAY [1.._MCCall.c_BufferDepthOutput] OF L_TS2P_FlexCamHighOut;
	_ASCPARCORE : ARRAY [1.._MCCall.c_BufferDepthInput] OF L_TS2P_scPar_FlexCamHigh;
	_ASCACCESSPOINTSCORE : ARRAY [1.._MCCall.c_BufferDepthInput] OF L_TS2P_scAP_FlexCamHigh;
	_ASCSIGNALFLOWCORE : ARRAY [1.._MCCall.c_BufferDepthOutput] OF L_TS2P_scSF_FlexCamHigh;
	_SCINPUTVISU : L_TS2P_FlexCamHighIn;
	_PSCINPUTVISU : POINTER TO L_TS2P_FlexCamHighIn := ADR(_scInputVisu);
	_PSCOUTPUTVISU : POINTER TO L_TS2P_FlexCamHighOut := ADR(_ascOutput[1]);
	_PSCDATAVISU : POINTER TO L_TS2P_scData_TM_FlexCam := ADR(scData_int);
	_PSCPARVISU : POINTER TO L_TS2P_scPar_FlexCamHigh := ADR(scPar_int);
	_PSCAPVISU : POINTER TO L_TS2P_scAP_FlexCamHigh;
	_PSCSFVISU : POINTER TO L_TS2P_scSF_FlexCamHigh;
	ITFBASICMOTIONBASE : L_TB2P.L_TB2P_IBasicMotionBase;
	ITFFLEXCAMEXTENSION : L_TS2P_IFlexCam;
	ITFITECHMODULEINTERNAL : L_TB2P_ITechModuleInternal;
	LRJERKDEC : LREAL;
	LRJOGGINGJERKDEC : LREAL;
	REMAININGTIMEOFPROFILE : LREAL;
	REMAININGTIMEOFPROFILEAVAILABLE : BOOL;
END_VAR
END_FUNCTION_BLOCK

METHOD CALL_ABC
VAR_INPUT
	ITFTECHMODULE : L_TB2P.L_TB2P_IBasicMotionBase;
	XQSPAPPLICATION : BOOL;
	XHALT : BOOL;
	XABORT : BOOL;
	XHOMEEXECUTE : BOOL;
	XJOGPOS : BOOL;
	XJOGNEG : BOOL;
	XFINISHPOSITIONING : BOOL;
	XMOVEVELEXECUTE : BOOL;
	XMOVEABSEXECUTE : BOOL;
	XMOVERELEXECUTE : BOOL;
	XENABLEOPERATION : BOOL;
	XRESETERROR : BOOL;
	XENABLEPOSITIVE : BOOL;
	XENABLENEGATIVE : BOOL;
	XDISABLESWLIMIT : BOOL;
	LROVERRIDE : LREAL;
	LROVERRIDEACC : LREAL;
	LROVERRIDEJERK : LREAL;
	XRESETHOMEPOSITION : BOOL;
	XCONTINUOUSUPDATE : BOOL;
	LRPOS_DIST : LREAL;
	LRVEL : LREAL;
	LRACC : LREAL;
	LRDEC : LREAL;
	LRJERK : LREAL;
	EDIRECTION : L_TB2P.MC_DIRECTION;
	SCHOMEEXTTP : L_TB2P.MC_TRIGGER_REF;
	XHOMEABSSWITCH : BOOL;
	XSPECIALABORTBEHAVIOR : BOOL;
	LRABORTDEC : LREAL;
	LRABORTJERK : LREAL;
END_VAR
VAR_OUTPUT
	XERROR : BOOL;
	EERRORID : L_TB2P.L_IE1P_Error;
	XFUNBUSY : BOOL;
	XFUNDONE : BOOL;
	XFUNCOMMANDABORTED : BOOL;
	EFUNSTATEACT : L_TB2P.L_MC1P_ABC_State;
	ECONTROLMODE : L_TB2P.L_MC1P_ControlMode;
	XISHOMED : BOOL;
	XHWLIMITSWITCHNEG : BOOL;
	XHWLIMITSWITCHPOS : BOOL;
	XSWLIMITENABLED : BOOL;
	XSWLIMITSWITCHNEG : BOOL;
	XSWLIMITSWITCHPOS : BOOL;
	EAXISTYPE : L_TB2P.L_MC1P_DriveType;
	EAXISSTATE : L_TB2P.L_MC1P_AXIS_STATE;
	XSTOACTIVE : BOOL;
	XREADYFOROPERATION : BOOL;
	XOPERATIONENABLED : BOOL;
	XREADYFORMOTION : BOOL;
	XAXISWARNING : BOOL;
	XAXISERROR : BOOL;
	EAXISERRORID : L_TB2P.L_IE1P_Error;
	XDRIVEWARNING : BOOL;
	XDRIVEERROR : BOOL;
	DWDRIVEERRORID : DWORD;
	LRACTPOS : LREAL;
	LRACTVEL : LREAL;
	LRSETPOSOUT : LREAL;
	LRSETVELOUT : LREAL;
	LRACTFOLLOWINGERROR : LREAL;
	XINPOSITION : BOOL;
	XSTANDSTILLSETVELOCITY : BOOL;
	XSTANDSTILLACTVELOCITY : BOOL;
	XCONSTANTVELOCITY : BOOL;
	XACCELERATING : BOOL;
	XDECELERATING : BOOL;
	XDIRECTIONPOSITIVE : BOOL;
	XDIRECTIONNEGATIVE : BOOL;
	XAXISAVAILABLE : BOOL;
END_VAR
VAR_IN_OUT
	AXIS : AXIS_REF;
END_VAR
END_METHOD

METHOD GET_PAP : POINTER TO L_TB2P_scAP_TM_MotionControl
END_METHOD

METHOD GET_PDATA : POINTER TO L_TS2P_scData_TM_FlexCam
END_METHOD

METHOD GET_PDATASP : POINTER TO L_TS2P_scData_TM_FlexCam
END_METHOD

METHOD GET_PPAR : POINTER TO L_TB2P.L_TB2P_scPar_TM_MotionControl
END_METHOD

METHOD GET_PSF : POINTER TO L_TB2P_scSF_TM_MotionControl
END_METHOD

METHOD CAM
VAR_INPUT
	ITFTECHMODULE : L_TS2P_IFlexCam;
	XENABLE : BOOL;
	XSYNCCAM : BOOL;
	SCCAMTABLE : L_MC2P.MC_CAM_REF;
	LRCYCMASTERPOS : LREAL;
	LRCYCMASTERVEL : LREAL;
	LRCYCMASTERACC : LREAL;
	LRSLAVEPOS : LREAL;
	LRSLAVEVEL : LREAL;
	LRSLAVEACC : LREAL;
	EOFFSETMODEMASTER : L_TS2P_OffsetMode := L_TS2P_OffsetMode.x_zero;
	ESCALINGMODEMASTER : L_TS2P_ScalingMode := L_TS2P_ScalingMode.x_zero;
	EOFFSETMODESLAVE : L_TS2P_OffsetMode := L_TS2P_OffsetMode.x_zero;
	ESCALINGMODESLAVE : L_TS2P_ScalingMode := L_TS2P_ScalingMode.x_zero;
	LRSETOFFSETMASTER : LREAL;
	LRSETOFFSETSLAVE : LREAL;
	LRSETSCALINGMASTER : LREAL;
	LRSETSCALINGSLAVE : LREAL;
	LRPROFGENMASTERVEL : LREAL;
	LRPROFGENMASTERACC : LREAL;
	LRPROFGENMASTERDEC : LREAL;
	LRPROFGENMASTERJERK : LREAL;
	LRPROFGENSLAVEVEL : LREAL;
	LRPROFGENSLAVEACC : LREAL;
	LRPROFGENSLAVEDEC : LREAL;
	LRPROFGENSLAVEJERK : LREAL;
	XPERIODIC : BOOL;
	XCAMCHANGEINSTANT : BOOL;
	XMASTERABSOLUTE : BOOL;
	XSLAVEABSOLUTE : BOOL;
END_VAR
VAR_OUTPUT
	XERROR : BOOL;
	EERRORID : L_IE1P.L_IE1P_Error;
	LRSETPOSOUT : LREAL;
	LRSETVELOUT : LREAL;
	LRSETACCOUT : LREAL;
	LRSETXPOSOUT : LREAL;
	LRSETXVELOUT : LREAL;
	LRSETXACCOUT : LREAL;
	LRSETYPOSOUT : LREAL;
	LRSETYVELOUT : LREAL;
	LRSETYACCOUT : LREAL;
	XENDOFPROFILE : BOOL;
	LRSETOFFSETMASTEROUT : LREAL;
	LRSETOFFSETSLAVEOUT : LREAL;
	LRCONVERTMASTERTOXPOS : LREAL;
	LRCAMPROFILERPOSOUT : LREAL;
	LRCONVERTYTOSLAVEPOS : LREAL;
	XDONE : BOOL;
	XBUSY : BOOL;
END_VAR
END_METHOD

METHOD CAMSEQUENCER
VAR_INPUT
	ITFTECHMODULE : L_TS2P_IFlexCam;
	XENABLE : BOOL;
	XCAMSEQUENCER : BOOL;
	XENDOFPROFILEIN : BOOL;
	CAMTABLE1 : L_MC2P.MC_CAM_REF;
	CAMTABLE2 : L_MC2P.MC_CAM_REF;
	CAMTABLE3 : L_MC2P.MC_CAM_REF;
	CAMTABLE4 : L_MC2P.MC_CAM_REF;
	XCAMCHANGEINSTANT : BOOL;
	XLOADCAMTABLE : BOOL;
	WSETCAMTABLE : WORD;
	EMODE : L_TS2P_CamSequenceMode := L_TS2P_CamSequenceMode.CyclicCam1;
END_VAR
VAR_OUTPUT
	XERROR : BOOL;
	EERRORID : L_IE1P_Error;
	CAMTABLEOUT : L_MC2P.MC_CAM_REF;
	XCAMTABLEVALID : BOOL;
END_VAR
END_METHOD

METHOD CLUTCH
VAR_INPUT
	ITFTECHMODULE : L_TS2P_IFlexCam;
	XENABLE : BOOL;
	XCLUTCHCLOSE : BOOL;
	ECLUTCHINMODE : L_TS2P_ClutchInMode;
	ECLUTCHOUTMODE : L_TS2P_ClutchOutMode;
	EALLOWEDDIRECTION : L_TB2P_AllowedDirection;
	LRCLUTCHINDIST : LREAL;
	LRCLUTCHOUTDIST : LREAL;
	LRCLUTCHOUTPOSITION : LREAL;
	LRCYCLICMASTERPOS : LREAL;
	LRCYCLICMASTERVEL : LREAL;
	LRCYCLICMASTERACC : LREAL;
	LRCYCLICAXISPOS : LREAL;
	LRCYCLICAXISVEL : LREAL;
	LRCYCLICAXISACC : LREAL;
	ETRAVERSINGRANGE : L_MC1P_TraversingRange;
	LRCYCLELENGTH : LREAL;
END_VAR
VAR_OUTPUT
	XERROR : BOOL;
	EERRORID : L_IE1P.L_IE1P_Error;
	XBUSY : BOOL;
	XDONE : BOOL;
	XSYNCHRONISED : BOOL;
	XACCDECSYNC : BOOL;
	LRSETPOSOUT : LREAL;
	LRSETVELOUT : LREAL;
	LRSETACCOUT : LREAL;
END_VAR
END_METHOD

METHOD HALT : BOOL
VAR_INPUT
	ITFTECHMODULE : L_TS2P_IFlexCam;
	XEXECUTE : BOOL;
	LRDEC : LREAL := 100;
	LRJERK : LREAL := 0;
END_VAR
VAR_OUTPUT
	XBUSY : BOOL;
	XDONE : BOOL;
	XCOMMANDABORTED : BOOL;
END_VAR
VAR_IN_OUT
	AXIS : AXIS_REF;
END_VAR
END_METHOD

METHOD MOVETOPARKPOS : BOOL
VAR_INPUT
	ITFTECHMODULE : L_TS2P_IFlexCam;
	XEXECUTEMOVETOPARKPOS : BOOL;
	EMOVETOPARKPOSMODE : L_TS2P_CamStopMode;
	LRPARKPOSITION : LREAL := 180;
	EPOSITIONINGDIRECTION : L_TS2P_SyncDirection := L_TS2P_SyncDirection.PositiveDirection;
	LRPOSITIONINGVEL : LREAL := 10;
	LRPOSITIONINGACC : LREAL := 100;
	LRPOSITIONINGDEC : LREAL := 100;
	LRJERK : LREAL := 0;
END_VAR
VAR_OUTPUT
	XBUSY : BOOL;
	XDONE : BOOL;
	XCOMMANDABORTED : BOOL;
END_VAR
VAR_IN_OUT
	AXIS : AXIS_REF;
END_VAR
END_METHOD

METHOD POSITIONFOLLOWER
VAR_INPUT
	ITFTECHMODULE : L_TS2P_IFlexCam;
	XENABLE : BOOL;
	LRPOSITION : LREAL;
	LRVELOCITY : LREAL;
	LRACCELERATION : LREAL;
	ESETVALUEMODE : L_MC1P_SetValueMode;
END_VAR
VAR_OUTPUT
	XERROR : BOOL;
	EERRORID : L_IE1P.L_IE1P_Error;
	XBUSY : BOOL;
END_VAR
END_METHOD

METHOD SYNCIN
VAR_INPUT
	ITFTECHMODULE : L_TS2P_IFlexCam;
	XENABLE : BOOL;
	XSYNCIN : BOOL;
	XSYNCPOSRESTORE : BOOL;
	ESYNCMODE : L_TS2P_SyncInMode;
	ESYNCDIRECTION : L_TS2P_SyncDirection;
	LRSYNCVEL : LREAL;
	LRSYNCACC : LREAL;
	LRSYNCDEC : LREAL;
	LRSYNCJERK : LREAL;
	LRPARKPOSITION : LREAL;
	LRCYCLICMASTERPOS : LREAL;
	LRCYCLICMASTERVEL : LREAL;
	LRCYCLICMASTERACC : LREAL;
	LRCYCLICAXISPOS : LREAL;
	LRCYCLICAXISVEL : LREAL;
	LRCYCLICAXISACC : LREAL;
END_VAR
VAR_OUTPUT
	XERROR : BOOL;
	EERRORID : L_IE1P.L_IE1P_Error;
	XBUSY : BOOL;
	XDONE : BOOL;
	XSYNCHRONISED : BOOL;
	XACCDECSYNC : BOOL;
	LRSETPOSOUT : LREAL;
	LRSETVELOUT : LREAL;
	LRSETACCOUT : LREAL;
	LROFFSETSYNCPOS : LREAL;
END_VAR
VAR_IN_OUT
	AXIS : AXIS_REF;
END_VAR
END_METHOD

METHOD REQUESTINTERFACE : BOOL
VAR_INPUT
	ID : DINT;
	PITFUNKNOWN : POINTER TO L_UBUP.L_UBUP_IUnknown;
END_VAR
END_METHOD

METHOD CALLFUNCTION
VAR_INPUT
	UIINPUTDATAIDX : UINT;
	UIOUTPUTDATAIDX : UINT;
END_VAR
END_METHOD

METHOD COPYINPUTS : BOOL
VAR_INPUT
	IDX : WORD;
END_VAR
END_METHOD

METHOD COPYOUTPUTS : BOOL
VAR_INPUT
	IDX : WORD;
END_VAR
END_METHOD

METHOD FUNCTIONWASCALLEDTWICE : BOOL
VAR_INPUT
	IDX : WORD;
END_VAR
END_METHOD

METHOD HANDLESTANDARDCALL : BOOL
END_METHOD

METHOD SYNCOUTPUTS
VAR_INPUT
	UICOPYOUTPUTFROMIDX : UINT;
	UICOPYOUTPUTTOIDX : UINT;
END_VAR
END_METHOD

METHOD FB_INIT : BOOL
VAR_INPUT
	BINITRETAINS : BOOL;
	BINCOPYCODE : BOOL;
END_VAR
END_METHOD

METHOD CALL_INTERNALCTRL
END_METHOD

METHOD GET_INTERNCAMTABLE : MC_CAM_REF
END_METHOD

METHOD GET_LRCAMXEND : LREAL
END_METHOD

METHOD GET_LRCAMXSTART : LREAL
END_METHOD

METHOD GET_LRCAMYEND : LREAL
END_METHOD

METHOD GET_LRCAMYSTART : LREAL
END_METHOD

METHOD GET_STCAMNAME : STRING
END_METHOD

METHOD GET_XCOMMUNICATION : BOOL
END_METHOD

(* ---- L_TS2P_FLEXCAMSTATE.pou ---- *)
FUNCTION_BLOCK L_TS2P_FLEXCAMSTATE EXTENDS L_TB2P_TechModuleBase
VAR_INPUT
	XENABLE : BOOL;
	XENABLEOPERATION : BOOL;
	XRESETERROR : BOOL;
	XQSPAPPLICATION : BOOL;
	XABORT : BOOL;
	XJOGPOS : BOOL;
	XJOGNEG : BOOL;
	XHOMEEXECUTE : BOOL;
	LROVERRIDE : LREAL := 1;
	SCCTRLBASICMOTION : L_TB2P_scCtrlBasicMotion;
	SCPAR : L_TS2P_scPar_FlexCamState;
	SCACCESSPOINTS : L_TS2P_scAP_FlexCamState;
	MASTERVALUES : L_MC1P_IAXIS_REF_MASTERVALUES;
	XSYNCIN : BOOL;
	XCAMCHANGEINSTANT : BOOL;
	LRSETOFFSETPOSX : LREAL;
	LRSETOFFSETPOSY : LREAL;
	LRSETSCALINGX : LREAL := 1;
	LRSETSCALINGY : LREAL := 1;
	CAMTABLE1 : MC_CAM_REF;
	CAMTABLE2 : MC_CAM_REF;
	CAMTABLE3 : MC_CAM_REF;
	CAMTABLE4 : MC_CAM_REF;
	WSETCAMTABLE : WORD := 1;
	XCAMSEQUENCER : BOOL;
END_VAR
VAR_OUTPUT
	XREADYFOROPERATION : BOOL;
	XOPERATIONENABLED : BOOL;
	XREADYFORMOTION : BOOL;
	XERROR : BOOL;
	XWARNING : BOOL;
	EERRORID : L_IE1P_Error;
	XSTOACTIVE : BOOL;
	XQSPACTIVE : BOOL;
	XABORTBUSY : BOOL;
	XABORTDONE : BOOL;
	XJOGGINGBUSY : BOOL;
	XHOMINGBUSY : BOOL;
	XHOMINGDONE : BOOL;
	XISHOMED : BOOL;
	ETMSTATE : L_TB2P_States := L_TB2P_States.DISABLED;
	SCSTATUSBASICMOTION : L_TB2P_scStatusBasicMotion;
	LRACTVEL : LREAL;
	LRSETVELOUT : LREAL;
	LRACTPOS : LREAL;
	LRSETPOSOUT : LREAL;
	LRACTFOLLOWINGERROR : LREAL;
	SCSIGNALFLOW : L_TS2P_scSF_FlexCamState;
	XSYNCHRONISED : BOOL;
	XACCDECSYNC : BOOL;
	XCAMMINGBUSY : BOOL;
	XENDOFPROFILE : BOOL;
	LROFFSETPOSX : LREAL;
	LROFFSETPOSY : LREAL;
	WACTIVECAMTABLE : WORD;
	XCAMSEQUENCERACTIVE : BOOL;
END_VAR
VAR_IN_OUT
	AXIS : AXIS_REF;
END_VAR
VAR
	TM_INT : L_TS2P_TM_FlexCamState := STRUCT(ModuleHandler := ModuleHandler);
	SCPAR_INT : L_TS2P_scPar_FlexCamState;
	_UICALLMFUNIDXINPUT : UINT := 1;
	_UICALLMFUNIDXOUTPUT : UINT := 1;
	_MCCALL : L_UM1P_MCCall;
	_ASCINPUT : ARRAY [1.._MCCall.c_BufferDepthInput] OF L_TS2P_FlexCamStateIn;
	_ASCOUTPUT : ARRAY [1.._MCCall.c_BufferDepthOutput] OF L_TS2P_FlexCamStateOut;
	_ASCPARCORE : ARRAY [1.._MCCall.c_BufferDepthInput] OF L_TS2P_scPar_FlexCamState;
	_ASCACCESSPOINTSCORE : ARRAY [1.._MCCall.c_BufferDepthInput] OF L_TS2P_scAp_FlexCamState;
	_ASCSIGNALFLOWCORE : ARRAY [1.._MCCall.c_BufferDepthOutput] OF L_TS2P_scSF_FlexCamState;
	_SCINPUTVISU : L_TS2P_FlexCamStateIn;
	_PSCINPUTVISU : POINTER TO L_TS2P_FlexCamStateIn := ADR(_scInputVisu);
	_PSCOUTPUTVISU : POINTER TO L_TS2P_FlexCamStateOut := ADR(_ascOutput[1]);
	_PSCPARVISU : POINTER TO L_TS2P_scPar_FlexCamState := ADR(scPar_int);
	ITFITECHMODULEINTERNAL : L_TB2P_ITechModuleInternal;
	LRJERKDEC : LREAL;
	LRJOGGINGJERKDEC : LREAL;
	REMAININGTIMEOFPROFILE : LREAL;
	REMAININGTIMEOFPROFILEAVAILABLE : BOOL;
END_VAR
END_FUNCTION_BLOCK

METHOD GET_INTERNCAMTABLE : MC_CAM_REF
END_METHOD

METHOD GET_LRCAMXEND : LREAL
END_METHOD

METHOD GET_LRCAMXSTART : LREAL
END_METHOD

METHOD GET_LRCAMYEND : LREAL
END_METHOD

METHOD GET_LRCAMYSTART : LREAL
END_METHOD

METHOD GET_STCAMNAME : STRING
END_METHOD

METHOD GET_XCOMMUNICATION : BOOL
END_METHOD

METHOD GET_PAP : POINTER TO L_TB2P_scAP_TM_MotionControl
END_METHOD

METHOD GET_PPAR : POINTER TO L_TB2P_scPar_TM_MotionControl
END_METHOD

METHOD GET_PSF : POINTER TO L_TB2P_scSF_TM_MotionControl
END_METHOD

METHOD CALLFUNCTION
VAR_INPUT
	UIINPUTDATAIDX : UINT;
	UIOUTPUTDATAIDX : UINT;
END_VAR
END_METHOD

METHOD COPYINPUTS : BOOL
VAR_INPUT
	IDX : WORD;
END_VAR
END_METHOD

METHOD COPYOUTPUTS : BOOL
VAR_INPUT
	IDX : WORD;
END_VAR
END_METHOD

METHOD FUNCTIONWASCALLEDTWICE : BOOL
VAR_INPUT
	IDX : WORD;
END_VAR
END_METHOD

METHOD HANDLESTANDARDCALL : BOOL
END_METHOD

METHOD SYNCOUTPUTS
VAR_INPUT
	UICOPYOUTPUTFROMIDX : UINT;
	UICOPYOUTPUTTOIDX : UINT;
END_VAR
END_METHOD

METHOD CALL_INTERNALCTRL
END_METHOD

(* ---- L_TS2P_FLYINGSAWSTATE.pou ---- *)
FUNCTION_BLOCK L_TS2P_FLYINGSAWSTATE EXTENDS L_TB2P_TechModuleBase
VAR_INPUT
	XUSEORIGINAL : BOOL;
	XENABLE : BOOL;
	XENABLEOPERATION : BOOL;
	XRESETERROR : BOOL;
	XQSPAPPLICATION : BOOL;
	XABORT : BOOL;
	XJOGPOS : BOOL;
	XJOGNEG : BOOL;
	XHOMEEXECUTE : BOOL;
	LROVERRIDE : LREAL := 1;
	SCCTRLBASICMOTION : L_TB2P_scCtrlBasicMotion;
	SCPAR : L_TS2P_scPar_FlyingSawState;
	SCACCESSPOINTS : L_TS2P_scAP_FlyingSawState;
	MASTERVALUES : L_MC1P_IAXIS_REF_MASTERVALUES;
	XSTARTFLYINGSAW : BOOL;
	XSYNCININSTANT : BOOL;
	XEXECUTENEXTCUT : BOOL;
	XEXECUTEGAP : BOOL;
	XSETCUTTINGLENGTHINSTANT : BOOL;
	LRCUTTINGLENGTH : LREAL;
	LRSYNCOVERRIDE : LREAL := 1;
	XSETMATERIALCOUNTER : BOOL;
	XMOVETOPARKPOS : BOOL;
	XRESUMETARGETPOS : BOOL;
	XRESETMARKSTACK : BOOL;
	SCTPRECDATA_MARKSENSOR : L_MC1P.L_MC1P_TpReceiveData;
END_VAR
VAR_OUTPUT
	XREADYFOROPERATION : BOOL;
	XOPERATIONENABLED : BOOL;
	XREADYFORMOTION : BOOL;
	XERROR : BOOL;
	XWARNING : BOOL;
	EERRORID : L_IE1P_Error;
	XSTOACTIVE : BOOL;
	XQSPACTIVE : BOOL;
	XABORTBUSY : BOOL;
	XABORTDONE : BOOL;
	XJOGGINGBUSY : BOOL;
	XHOMINGBUSY : BOOL;
	XHOMINGDONE : BOOL;
	XISHOMED : BOOL;
	ETMSTATE : L_TB2P_States := L_TB2P_States.DISABLED;
	SCSTATUSBASICMOTION : L_TB2P_scStatusBasicMotion;
	LRACTVEL : LREAL;
	LRSETVELOUT : LREAL;
	LRACTPOS : LREAL;
	LRSETPOSOUT : LREAL;
	LRACTFOLLOWINGERROR : LREAL;
	SCSIGNALFLOW : L_TS2P_scSF_FlyingSawState;
	XSYNCHRONISED : BOOL;
	XACCDECSYNC : BOOL;
	XINPOSITION : BOOL;
	XPOSITIONING : BOOL;
	LRMATERIALCOUNTER : LREAL;
	LRTARGETPOS : LREAL;
	LRCUTGAP : LREAL;
	LRACTIVECUTTINGLENGTH : LREAL;
	WMARKSINSTACK : WORD;
END_VAR
VAR_IN_OUT
	AXIS : AXIS_REF;
END_VAR
VAR
	XINTERNALCONTROLACTIVE_OLD : BOOL;
	XUSEORIGINAL_OLD : BOOL;
	ITFCONNECTORFLYINGSAW : L_TS2P_IConnectorFlyingSaw;
	TM_INT : L_TS2M_TM_FlyingSawState;
	SCPAR_INT : L_TS2P_scPar_FlyingSawState;
	_SCDATA_INT : L_TS2M_scData_FlyingSawState;
	_SCFMDATA_INT : L_TS2M_scData_FM_FlyingSaw;
	_UICALLMFUNIDXINPUT : UINT := 1;
	_UICALLMFUNIDXOUTPUT : UINT := 1;
	_MCCALL : L_UM1P_MCCall;
	_ASCINPUT : ARRAY [1.._MCCall.c_BufferDepthInput] OF L_TS2P_FlyingSawStateIn;
	_ASCOUTPUT : ARRAY [1.._MCCall.c_BufferDepthOutput] OF L_TS2P_FlyingSawStateOut;
	_ASCPARCORE : ARRAY [1.._MCCall.c_BufferDepthInput] OF L_TS2P_scPar_FlyingSawState;
	_ASCACCESSPOINTSCORE : ARRAY [1.._MCCall.c_BufferDepthInput] OF L_TS2P_scAP_FlyingSawState;
	_ASCSIGNALFLOWCORE : ARRAY [1.._MCCall.c_BufferDepthOutput] OF L_TS2P_scSF_FlyingSawState;
	_ASCDATACORE : ARRAY [1.._MCCall.c_BufferDepthInput] OF L_TS2M_scData_FlyingSawState;
	_ASCDATAFMCORE : ARRAY [1.._MCCall.c_BufferDepthInput] OF L_TS2M_scData_FM_FlyingSaw;
	_SCINPUTVISU : L_TS2P_FlyingSawStateIn;
	_PSCINPUTVISU : POINTER TO L_TS2P_FlyingSawStateIn := ADR(_scInputVisu);
	_PSCOUTPUTVISU : POINTER TO L_TS2P_FlyingSawStateOut := ADR(_ascOutput[1]);
	_PSCPARVISU : POINTER TO L_TS2P_scPar_FlyingSawState := ADR(scPar_int);
	_PSCDATAVISU : POINTER TO L_TS2M_scData_FlyingSawState := ADR(_scData_int);
	_PSCFMDATAVISU : POINTER TO L_TS2M_scData_FM_FlyingSaw := ADR(_scFMData_int);
	_PSCFMSFVISU : POINTER TO L_TS2P_scSF_FlyingSawState;
	ITFBASICMOTIONBASE : L_TB2P.L_TB2P_IBasicMotionBase;
	ITFFLYINGSAWPROCESSINGEXTENSION : L_TS2P_IFlyingSawProcessing;
	ITFITECHMODULEINTERNAL : L_TB2P_ITechModuleInternal;
	LRJERKDEC : LREAL;
	LRJOGGINGJERKDEC : LREAL;
	REMAININGTIMEOFPROFILE : LREAL;
	REMAININGTIMEOFPROFILEAVAILABLE : BOOL;
END_VAR
END_FUNCTION_BLOCK

METHOD CALL_ABC
VAR_INPUT
	ITFTECHMODULE : L_TB2P.L_TB2P_IBasicMotionBase;
	XQSPAPPLICATION : BOOL;
	XHALT : BOOL;
	XABORT : BOOL;
	XHOMEEXECUTE : BOOL;
	XJOGPOS : BOOL;
	XJOGNEG : BOOL;
	XFINISHPOSITIONING : BOOL;
	XMOVEVELEXECUTE : BOOL;
	XMOVEABSEXECUTE : BOOL;
	XMOVERELEXECUTE : BOOL;
	XENABLEOPERATION : BOOL;
	XRESETERROR : BOOL;
	XENABLEPOSITIVE : BOOL;
	XENABLENEGATIVE : BOOL;
	XDISABLESWLIMIT : BOOL;
	LROVERRIDE : LREAL;
	LROVERRIDEACC : LREAL;
	LROVERRIDEJERK : LREAL;
	XRESETHOMEPOSITION : BOOL;
	XCONTINUOUSUPDATE : BOOL;
	LRPOS_DIST : LREAL;
	LRVEL : LREAL;
	LRACC : LREAL;
	LRDEC : LREAL;
	LRJERK : LREAL;
	EDIRECTION : L_TB2P.MC_DIRECTION;
	SCHOMEEXTTP : L_TB2P.MC_TRIGGER_REF;
	XHOMEABSSWITCH : BOOL;
	XSPECIALABORTBEHAVIOR : BOOL;
	LRABORTDEC : LREAL;
	LRABORTJERK : LREAL;
END_VAR
VAR_OUTPUT
	XERROR : BOOL;
	EERRORID : L_TB2P.L_IE1P_Error;
	XFUNBUSY : BOOL;
	XFUNDONE : BOOL;
	XFUNCOMMANDABORTED : BOOL;
	EFUNSTATEACT : L_TB2P.L_MC1P_ABC_State;
	ECONTROLMODE : L_TB2P.L_MC1P_ControlMode;
	XISHOMED : BOOL;
	XHWLIMITSWITCHNEG : BOOL;
	XHWLIMITSWITCHPOS : BOOL;
	XSWLIMITENABLED : BOOL;
	XSWLIMITSWITCHNEG : BOOL;
	XSWLIMITSWITCHPOS : BOOL;
	EAXISTYPE : L_TB2P.L_MC1P_DriveType;
	EAXISSTATE : L_TB2P.L_MC1P_AXIS_STATE;
	XSTOACTIVE : BOOL;
	XREADYFOROPERATION : BOOL;
	XOPERATIONENABLED : BOOL;
	XREADYFORMOTION : BOOL;
	XAXISWARNING : BOOL;
	XAXISERROR : BOOL;
	EAXISERRORID : L_TB2P.L_IE1P_Error;
	XDRIVEWARNING : BOOL;
	XDRIVEERROR : BOOL;
	DWDRIVEERRORID : DWORD;
	LRACTPOS : LREAL;
	LRACTVEL : LREAL;
	LRSETPOSOUT : LREAL;
	LRSETVELOUT : LREAL;
	LRACTFOLLOWINGERROR : LREAL;
	XINPOSITION : BOOL;
	XSTANDSTILLSETVELOCITY : BOOL;
	XSTANDSTILLACTVELOCITY : BOOL;
	XCONSTANTVELOCITY : BOOL;
	XACCELERATING : BOOL;
	XDECELERATING : BOOL;
	XDIRECTIONPOSITIVE : BOOL;
	XDIRECTIONNEGATIVE : BOOL;
	XAXISAVAILABLE : BOOL;
END_VAR
VAR_IN_OUT
	AXIS : AXIS_REF;
END_VAR
END_METHOD

METHOD GET_PAP : POINTER TO L_TB2P_scAP_TM_MotionControl
END_METHOD

METHOD GET_PDATA : POINTER TO L_TS2M_scData_FlyingSawState
END_METHOD

METHOD GET_PFMDATA : POINTER TO L_TS2M_scData_FM_FlyingSaw
END_METHOD

METHOD GET_PPAR : POINTER TO L_TB2P_scPar_TM_MotionControl
END_METHOD

METHOD GET_PSF : POINTER TO L_TB2P_scSF_TM_MotionControl
END_METHOD

METHOD CLUTCH
VAR_INPUT
	ITFTECHMODULE : L_TS2P_IFlyingSawProcessing;
	XENABLE : BOOL;
	XSYNCVEL : BOOL := FALSE;
	XSYNCPOS : BOOL;
	XSYNCOUTINSTANT : BOOL;
	LRSYNCVEL : LREAL := 10;
	LRSYNCACC : LREAL := 100;
	LRSYNCDEC : LREAL := 100;
	LRSYNCJERK : LREAL := 10000;
	LRCYCMASTERPOS : LREAL;
	LRCYCMASTERVEL : LREAL;
	LRCYCMASTERACC : LREAL;
	LRSETSLAVEPOS : LREAL;
	LRSETSLAVEVEL : LREAL;
	LRSETSLAVEACC : LREAL;
END_VAR
VAR_OUTPUT
	EERRORID : L_IE1P.L_IE1P_Error;
	XERROR : BOOL;
	XBUSY : BOOL;
	XDONE : BOOL;
	XACCDECSYNC : BOOL;
	XVELSYNCHRONISED : BOOL;
	XPOSSYNCHRONISED : BOOL;
	LRSETSLAVEPOSOUT : LREAL;
	LRSETSLAVEVELOUT : LREAL;
	LRSETSLAVEACCOUT : LREAL;
	XPROFILERESETTIMEVALID : BOOL;
	LRPROFILERESETTIME : LREAL;
END_VAR
END_METHOD

METHOD EXECUTEGAP
VAR_INPUT
	ITFTECHMODULE : L_TS2P_IFlyingSawProcessing;
	XENABLE : BOOL;
	LRSYNCVEL : LREAL := 10;
	LRSYNCACC : LREAL := 100;
	LRSYNCDEC : LREAL := 100;
	LRSYNCJERK : LREAL := 10000;
	XEXECUTEGAP : BOOL;
	XAUXEXECUTEGAP : BOOL := FALSE;
	LRCYCMASTERPOS : LREAL;
	LRCYCMASTERVEL : LREAL;
	LRCYCMASTERACC : LREAL;
	LRSETSLAVEPOS : LREAL;
	LRSETSLAVEVEL : LREAL;
	LRSETSLAVEACC : LREAL;
END_VAR
VAR_OUTPUT
	EERRORID : L_IE1P.L_IE1P_Error;
	XERROR : BOOL;
	XBUSY : BOOL;
	XDONE : BOOL;
	XACCDECSYNC : BOOL;
	XVELSYNCHRONISED : BOOL;
	XPOSSYNCHRONISED : BOOL;
	LRSETSLAVEPOSOUT : LREAL;
	LRSETSLAVEVELOUT : LREAL;
	LRSETSLAVEACCOUT : LREAL;
	XPROFILERESETTIMEVALID : BOOL;
	LRPROFILERESETTIME : LREAL;
END_VAR
END_METHOD

METHOD MARKSTACK_GETMARK
VAR_INPUT
	ITFTECHMODULE : L_TS2P_IFlyingSawProcessing;
	XENABLE : BOOL;
	XGETMARK : BOOL;
	XRESETGETMARK : BOOL;
	XRESETMARKSTACK : BOOL;
	LRCYCSETPOS : LREAL;
	LRCYCSETVEL : LREAL;
END_VAR
VAR_OUTPUT
	XMARKSTACKFULL : BOOL;
	XMARKSTACKEMPTY : BOOL;
	WMARKSINSTACK : WORD;
	XMARKVALID : BOOL;
	LRMARKPOSOUT : LREAL;
END_VAR
END_METHOD

METHOD MARKSTACK_SETMARK
VAR_INPUT
	ITFTECHMODULE : L_TS2P_IFlyingSawProcessing;
	XENABLE : BOOL;
	XSETMARK : BOOL;
	LRMARKPOS : LREAL;
	XRESETMARKSTACK : BOOL;
	LRCYCSETPOS : LREAL;
	LRCYCSETVEL : LREAL;
END_VAR
VAR_OUTPUT
	XMARKSTACKFULL : BOOL;
	XMARKSTACKEMPTY : BOOL;
	WMARKSINSTACK : WORD;
	XNEWMARKRECEIVED : BOOL;
END_VAR
END_METHOD

METHOD POSITIONING
VAR_INPUT
	ITFTECHMODULE : L_TS2P_IFlyingSawProcessing;
	XENABLE : BOOL;
	XMOVETOTARGETPOS : BOOL;
	LRTARGETPOS : LREAL;
	LRPOSITIONINGVEL : LREAL;
	LRPOSITIONINGACC : LREAL;
	LRPOSITIONINGDEC : LREAL;
	LRPOSITIONINGJERK : LREAL;
	LRSETSLAVEPOS : LREAL;
	LRSETSLAVEVEL : LREAL;
	LRSETSLAVEACC : LREAL;
	LRCORRECTTIMEBASE : LREAL := 0;
	LROVERRIDE : LREAL := 1.0;
END_VAR
VAR_OUTPUT
	EERRORID : L_IE1P.L_IE1P_Error;
	XERROR : BOOL;
	XBUSY : BOOL;
	XDONE : BOOL;
	XPOSITIONING : BOOL;
	XINPOSITION : BOOL;
	LRSETSLAVEPOSOUT : LREAL;
	LRSETSLAVEVELOUT : LREAL;
	LRSETSLAVEACCOUT : LREAL;
	XPROFILERESETTIMEVALID : BOOL;
	LRPROFILERESETTIME : LREAL;
END_VAR
END_METHOD

METHOD REQUESTINTERFACE : BOOL
VAR_INPUT
	ID : DINT;
	PITFUNKNOWN : POINTER TO L_UBUP.L_UBUP_IUnknown;
END_VAR
END_METHOD

METHOD CALLFUNCTION
VAR_INPUT
	UIINPUTDATAIDX : UINT;
	UIOUTPUTDATAIDX : UINT;
END_VAR
END_METHOD

METHOD COPYINPUTS : BOOL
VAR_INPUT
	IDX : WORD;
END_VAR
END_METHOD

METHOD COPYOUTPUTS : BOOL
VAR_INPUT
	IDX : WORD;
END_VAR
END_METHOD

METHOD FUNCTIONWASCALLEDTWICE : BOOL
VAR_INPUT
	IDX : WORD;
END_VAR
END_METHOD

METHOD HANDLESTANDARDCALL : BOOL
END_METHOD

METHOD SYNCOUTPUTS
VAR_INPUT
	UICOPYOUTPUTFROMIDX : UINT;
	UICOPYOUTPUTTOIDX : UINT;
END_VAR
END_METHOD

METHOD FB_INIT : BOOL
VAR_INPUT
	BINITRETAINS : BOOL;
	BINCOPYCODE : BOOL;
END_VAR
END_METHOD

METHOD CALL_INTERNALCTRL
END_METHOD

(* ---- L_TS2P_INVERTGEARFACTOR.pou ---- *)
FUNCTION_BLOCK L_TS2P_INVERTGEARFACTOR
VAR_INPUT
	XINVERTGEARFACTOR : BOOL;
	LRCYCLELENGTHX : LREAL := 1.0;
	LRCYCLELENGTHY : LREAL := 1.0;
	LRCOUPLINGX : LREAL := 1.0;
	LRCOUPLINGY : LREAL := 1.0;
	XDISABLETOLERANCEINVERTGEARFACTOR : BOOL;
	LRTOLERANCEINVERTGEARFACTOR : LREAL := 0;
END_VAR
VAR_OUTPUT
	XINVERTGEARFACTORACTIVE : BOOL;
	LRCYCLELENGTHX_OUT : LREAL;
	LRCYCLELENGTHY_OUT : LREAL;
	LRCOUPLINGX_OUT : LREAL;
	LRCOUPLINGY_OUT : LREAL;
	XWARNING : BOOL;
	EERRORID : L_IE1P_Error;
END_VAR
VAR_IN_OUT
	AXIS : AXIS_REF;
END_VAR
VAR
	XINWINDOW : BOOL;
END_VAR
END_FUNCTION_BLOCK

(* ---- L_TS2P_MARKQUEUE.pou ---- *)
FUNCTION_BLOCK L_TS2P_MARKQUEUE
VAR_INPUT
	XENABLE : BOOL;
	XLOADMARKPOS : BOOL;
	LRMARKPOS : LREAL;
	XGETNEXTMARK : BOOL;
	XRESETGETNEXTMARK : BOOL;
	XRESETMARKQUEUE : BOOL;
	LRCYCSETPOS : LREAL;
	LRCYCSETVEL : LREAL;
END_VAR
VAR_OUTPUT
	XQUEUEISFULL : BOOL;
	XQUEUEISEMPTY : BOOL;
	XNEWMARKRECEIVED : BOOL;
	WMARKSINQUEUE : WORD;
	XMARKVALID : BOOL;
	LRMARKPOSOUT : LREAL;
END_VAR
VAR
	FB_MB1P_STACK : L_MB1P_Stack;
	XTRACKMARK : BOOL;
	XENABLE_OLD : BOOL;
	XRESETMARKQUEUE_OLD : BOOL;
	XGETNEXTMARK_OLD : BOOL;
	XRESETGETNEXTMARK_OLD : BOOL;
	C_LRMATERIALCOUNTERCYCLELENGTH : LREAL := (16#4FFFFFFFFFFFFFFF * 1E-08);
END_VAR
END_FUNCTION_BLOCK

(* ---- L_TS2P_MARKSTACK.pou ---- *)
FUNCTION_BLOCK L_TS2P_MARKSTACK
VAR_INPUT
	XENABLE : BOOL;
	TPRECDATAIN : L_MC1P_TpReceiveData;
	LRACTVELMATERIAL : LREAL;
	LRACTPOSITIONTPAXIS : LREAL;
	LRCYCLELENGTHTPAXIS : LREAL;
	LRMARKSTACKLENGTH : LREAL;
	LRTASKCYCLE : LREAL;
END_VAR
VAR_OUTPUT
	TPRECDATAOUT : L_MC1P_TpReceiveData;
	XERROR : BOOL := FALSE;
	EERRORID : WORD;
	LRTPDIFFOUT : LREAL;
END_VAR
VAR
	ALRINTEGRATORSTARTPOS : ARRAY [1..64] OF LREAL := [64(0)];
	ALRLASTSCAN : ARRAY [1..64] OF LREAL := [64(0)];
	ALRDUMMY : ARRAY [1..64] OF LREAL := [64(0)];
	AXTPVALID : ARRAY [1..64] OF BOOL := [64(FALSE)];
	AXDUMMY : ARRAY [1..64] OF BOOL := [64(FALSE)];
	ADWACTTIMESTAMP : ARRAY [1..64] OF DWORD := [64(0)];
	ADWRECTIMESTAMP : ARRAY [1..64] OF DWORD := [64(0)];
	ADWDUMMY : ARRAY [1..64] OF DWORD := [64(0)];
	XREGISTERFULL : BOOL := FALSE;
	XINIT : BOOL := TRUE;
	WCOUNTER : WORD;
	WCOUNTERIN : WORD := 1;
	WCOUNTEROUT : WORD := 1;
	LRINTEGRATORPOS : LREAL := 0;
	LRCYCPOSDIFF : LREAL := 0;
	LRPOSTOREGISTEREND : LREAL := 0;
	XTPRECEIVEDINOLD : BOOL;
	LRMARKSTACKLENGTHOLD : LREAL;
	LRACTPOSITIONTPAXISCOMP : LREAL;
	LRACTTPPOSITIONOUT_INT : LREAL;
	DWDEADTIMESTACKOUT : DWORD;
	LRINTEGRATORLENGTH : LREAL := 10000000000.0;
END_VAR
END_FUNCTION_BLOCK

METHOD CALL_INITMARKSTACK
END_METHOD

(* ---- L_TS2P_MARKSTACKFLYINGSAW.pou ---- *)
FUNCTION_BLOCK L_TS2P_MARKSTACKFLYINGSAW
VAR
	FB_MB1P_STACK : L_MB1P_Stack_FlyingSaw;
	XTRACKMARK : BOOL;
	XMARKVALID_INT : BOOL;
	XENABLE_OLD : BOOL;
	XRESETMARKSTACK_OLD : BOOL;
	XGETMARK_OLD : BOOL;
	XSETMARK_OLD : BOOL;
	XRESETGETMARK_OLD : BOOL;
	C_LRMATERIALCOUNTERCYCLELENGTH : LREAL := (16#4FFFFFFFFFFFFFFF * 1E-08);
END_VAR
END_FUNCTION_BLOCK

METHOD DISABLE
END_METHOD

METHOD RESETMARKSTACK
END_METHOD

METHOD GETMARK
VAR_INPUT
	XENABLE : BOOL;
	XGETMARK : BOOL;
	XRESETGETMARK : BOOL;
	XRESETMARKSTACK : BOOL;
	LRCYCSETPOS : LREAL;
	LRCYCSETVEL : LREAL;
END_VAR
VAR_OUTPUT
	XMARKSTACKFULL : BOOL;
	XMARKSTACKEMPTY : BOOL;
	WMARKSINSTACK : WORD;
	XMARKVALID : BOOL;
	LRMARKPOSOUT : LREAL;
END_VAR
END_METHOD

METHOD SETMARK
VAR_INPUT
	XENABLE : BOOL;
	XSETMARK : BOOL;
	LRMARKPOS : LREAL;
	XRESETMARKSTACK : BOOL;
	LRCYCSETPOS : LREAL;
	LRCYCSETVEL : LREAL;
END_VAR
VAR_OUTPUT
	XMARKSTACKFULL : BOOL;
	XMARKSTACKEMPTY : BOOL;
	WMARKSINSTACK : WORD;
	XNEWMARKRECEIVED : BOOL;
END_VAR
END_METHOD

(* ---- L_TS2P_MARKWINDOWRELATIVE.pou ---- *)
FUNCTION_BLOCK L_TS2P_MARKWINDOWRELATIVE
VAR_INPUT
	XENABLE : BOOL;
	LRTPWINDOWSIZE : LREAL;
	LRSETOFFSETTPWINDOW : LREAL;
	LRCYCVEL : LREAL;
	TPRECDATAIN : L_MC1P_TpReceiveData;
	LRSTARTPOSITION : LREAL;
	LRCYCLELENGTH : LREAL;
	XTEACHMARKWINDOW : BOOL;
	DWMAXTPNOTDETECTED : DWORD;
	LRTASKCYCLE : LREAL;
END_VAR
VAR_OUTPUT
	TPRECDATAOUT : L_MC1P_TpReceiveData;
	XTPWINDOWOPEN : BOOL;
	XTPWINDOWOPENCOMP : BOOL;
	LRTPDELTAPOSCOMP : LREAL;
	XTPINWINDOW : BOOL;
	XTPNOTINWINDOW : BOOL;
	XTPNOTDETECTED : BOOL;
	XTPSENSORTEACHED : BOOL;
	XMAXTPNOTDETECTED : BOOL;
END_VAR
VAR
	LRMARKWINDOWINTEGRATOROLD : LREAL;
	XTPNOTDETECTEDINTERNAL : BOOL;
	LRLOWERWINDOW : LREAL;
	LRUPPERWINDOW : LREAL;
	XTEACHTPSENSOROLD : BOOL;
	DWMISSEDTPCOUNTER : DWORD;
	XTPISINWINDOW : BOOL;
	LRDEADTIMEPOSDIFF : LREAL;
	LRUPPERWINDOWCOMP : LREAL;
	XTPCOMPWINDOWOPEN : BOOL;
	XTPCOMPWINDOWOPENOLD : BOOL := FALSE;
	LRLOWERWINDOWCOMP : LREAL;
	XTPRECEIVEDOLD : BOOL;
	XTPRECEIVEDINTERNAL : BOOL;
	LRTPWINDOWSIZE_INT : LREAL;
	LRMARKWINDOWINTEGRATOR : LREAL := 0;
	LRDEADTIMETP : LREAL;
	LRACTUALTPPOSITION : LREAL;
END_VAR
END_FUNCTION_BLOCK

(* ---- L_TS2P_MASTERVALUECORRECTION.pou ---- *)
FUNCTION_BLOCK L_TS2P_MASTERVALUECORRECTION
VAR_INPUT
	XAXIS : POINTER TO L_MC1P_IAXIS_REF_MASTERVALUES;
	XENABLE : BOOL;
	XENABLECORRECTION : BOOL;
	XRESETERROR : BOOL;
	LRSETVELIN : LREAL;
	LRACTPOSITIONTOOL : LREAL;
	LRCYCLELENGTHTOOL : LREAL;
	TPRECDATA : L_MC1P_TpReceiveData;
	XLOADREGPOS : BOOL;
	LRLOADREGPOS : LREAL;
	LRSENSORTOOLDIST : LREAL;
	LRMARKDIST : LREAL;
	LRMAXCORRNEG : LREAL;
	LRMAXCORRPOS : LREAL;
	ESOURCEFORCORRWINDOW : L_TS2P_SourceForCorrWindow;
	LRUPPERCORRPOS : LREAL;
	LRLOWERCORRPOS : LREAL;
	DWGEARINGNUMERATORY : DWORD := 1;
	DWGEARINGDENOMINATORY : DWORD := 1;
	XSYNCHRONISED : BOOL;
	LRACTOFFSETMASTERIN : LREAL;
	LRACTOFFSETSLAVEIN : LREAL;
	XTEACHMARKWINDOW : BOOL;
	XENABLEMARKWINDOW : BOOL;
	LRMARKWINDOWSIZE : LREAL;
	LRSETOFFSETMARKWINDOW : LREAL;
	DWMAXNUMBERVIRTUALMARKS : DWORD;
	LRGEARFACTORCORRGAIN : LREAL;
	LRMAXGEARFACTORCORR : LREAL;
	XGEARFACTORCORR : BOOL;
	XGEARFACTORCORRHOLD : BOOL;
	XENABLETOOLCORRECTION : BOOL;
	LRTRANSMITCYCLESSETPOS : LREAL;
	DIDEADTIMECOMP : DINT;
	LRCORRVEL : LREAL;
	LRCORRACC : LREAL;
	LRCORRDEC : LREAL;
	LRCORRJERK : LREAL;
	ECORRMODE : L_TS2P_CorrectionMode;
	ECORRMODEOLD : L_TS2P_CorrectionMode;
END_VAR
VAR_OUTPUT
	CORRECTEDXAXIS : L_MC1P_IAXIS_REF_MASTERVALUES;
	LRACTVEL : LREAL;
	XERROR : BOOL;
	XWARNING : BOOL;
	EERRORID : WORD;
	XCORRLIMITED : BOOL;
	LRACTMARKERROR : LREAL;
	LRACTMARKDIST : LREAL;
	XINITDONE : BOOL;
	XCORRACTIVE : BOOL;
	XMARKRECEIVED : BOOL;
	LRSENSORACTPOS : LREAL;
	LRSENSORSETPOS : LREAL;
	XMARKWINDOWOPEN : BOOL;
	XMARKOUTOFWINDOW : BOOL;
	XMARKNOTDETECTED : BOOL;
	XMARKWINDOWTEACHED : BOOL;
	LRGEARFACTORCORR : LREAL;
	XGEARFACTORCORRLIMITED : BOOL;
	XCORRNEXTCYCLE : BOOL;
END_VAR
VAR_IN_OUT
	YAXIS : AXIS_REF;
END_VAR
VAR
	FB_L_TB2P_TP_CONVERTER : L_TB2P_TP_Converter;
	FB_L_TS2P_MARKWINDOWRELATIVE : L_TS2P_MarkWindowRelative;
	FB_L_TS2P_TPVIRTUALACTPOS : L_TS2P_TpVirtualActPos;
	FB_L_TS2P_MARKSTACK : L_TS2P_MarkStack;
	FB_L_MC1P_TPCALCDIFF : L_MC1P_TpCalcDiff;
	FB_L_TS2P_TPLIMITDIFF : L_TS2P_TpLimitDiff;
	FB_L_TS2P_DISTCORRECTIONWINDOW : L_TS2P_DistCorrectionWindow;
	FB_L_MC1P_SETAXISREFMASTERVALUES : L_MC1P_SetAxisRefMasterValues;
	FB_PROFILEGENERATOR : L_MC1P_ProfileGenerator;
	FB_INTEGRATOR : L_MC1P_IntegrateAxis;
	SCPROFILEPARAMETER : L_MC1P_ProfileParameter;
	FB_RAMPGENERATORGEARFACTOR : L_MC1P_RampGenerator;
	LRSENSORSETPOS_INT : LREAL;
	LRGEARINGFAKTOR : LREAL := 1.0;
	LRTPDIFFERENCE_INT : LREAL;
	XTPINWINDOW : BOOL;
	XVALUESTOREDTPCONVERTER : BOOL;
	XVALUESTOREDTPCONVERTEROLD : BOOL;
	XVALUESTOREDMARKWINDOW : BOOL;
	XVALUESTOREDMISSEDMARKS : BOOL;
	XVALUESTOREDMARKSTACK : BOOL;
	XVALUESTOREDCALCDIFF : BOOL;
	XVALUESTOREDLIMIT : BOOL;
	LRCORRRESIDUAL : LREAL;
	LRTPACTPOSITION_INT : LREAL;
	LRTPDIFFERENCELIM_INT : LREAL;
	LROFFSETPOSCTRL_INT : LREAL;
	LRCYCVELIN_INT : LREAL;
	LRSETCORRECTEDPOSOUT_INT : LREAL;
	LRMASTERSETPOSOLD_INT : LREAL;
	LRCORRPOSOUTOLD_INT : LREAL;
	LRVELOUT_INT : LREAL;
	XCORRACTIVE_INT : BOOL;
	XINIT : BOOL := TRUE;
	XTPCORRECTIONACTIVE : BOOL := FALSE;
	LRTPAXISSETPOS : LREAL;
	LRMARKDIST_INT : LREAL;
	XZERO : BOOL;
	XHOMINGDONE : BOOL;
	XSTARTREFERENCEACTIVE : BOOL;
	XHOMINGACTIVE : BOOL := FALSE;
	XMARKDISTCHANGED : BOOL;
	XENABLE_OLD : BOOL;
	XTPRECEIVEDOUT_INTOLD : BOOL;
	XSTARTFIRSTCORRECTION : BOOL;
	LRTPDIFFERENCELIM2_INT : LREAL;
	XCORRECTIONBUSYOLD : BOOL;
	LRTPACTPOSIN_OLD : LREAL;
	LRTPSETPOSIN_OLD : LREAL;
	LRTPAXISACTPOS_OLD : LREAL;
	LRCYCLELENGTH : LREAL;
	ICOUNTER : INT := 0;
	LRSETPOSITIONOLD : LREAL;
	LRCYCLELENGTHTP : LREAL;
	LRTPACTPOSITIONOLD : LREAL;
	XFIRSTTOUCHPROBE : BOOL := TRUE;
	LRSENSORTOOLDISTANCE_INT : LREAL;
	LRMARKSTACKLENGTH : LREAL;
	LRTPDIFFERENCELIMITOUT_INT : LREAL;
	XTPNOTDETECTED_INT : BOOL;
	XMAXTPNOTDETECTED : BOOL;
	LRGEARINGFAKTOROLD : LREAL;
	LRGEARFACTORINTEGRATOR : LREAL;
	LRGEARFACTORGAIN : LREAL := 1;
	LRGEARFACTORNUMERATORCORR : LREAL;
	LRGEARFACTORNUMERATORCORRLIMITED : LREAL;
	LRGEARFACTORDENOMINATOR : LREAL;
	LRGEARFACTORNUMERATOR : LREAL;
	LRTOTALSTACKDIFFERENCEOUT_INT : LREAL := 0;
	LCORRECTIONVELIN : LREAL;
	LRSETPOSCORROUT_OLD : LREAL;
	LRDELTAGEARFACTORCORR : LREAL;
	XTPSENSORTEACHEDOLD : BOOL;
	XTPSENSORTEACHEDATLASTMARK : BOOL;
	XCALCMARKDISTINITIALISED : BOOL;
	XTEACHTPSENSOROLD : BOOL;
	LRTPDEADTIMEDIFF : LREAL;
	XTPRECEIVEDOUTOLD_INT : BOOL;
	LRMARKDISTINTEGRATOR : LREAL;
	LRTPAXISCOMPFACTOR : LREAL;
	LRTPAXISDELAYCYCLE : LREAL;
	XENABLEOLD : BOOL;
	XTPRECEIVEDINOLD_INT : BOOL;
	TPRECDATAMARKWINDOW : L_MC1P_TpReceiveData;
	TPRECDATAMARKSTACK : L_MC1P_TpReceiveData;
	LRMASTERACTPOSITIONOLD_INT : LREAL;
	XFIRSTVALUESTORED : BOOL := FALSE;
	LRSETINTEGRATEDPOSITIONOLD : LREAL;
	XRESETERROROLD : BOOL;
	LRTPDIFF : LREAL;
	LRVELDIFF : LREAL;
	LRVELCOMP : LREAL;
	SETPOSITIONFORSYNCOLD : LREAL;
	LRMARKDISTOLD : LREAL;
END_VAR
END_FUNCTION_BLOCK

METHOD CALL_CALCACTMARKDIST
END_METHOD

METHOD CALL_CALCMARKERROR
END_METHOD

METHOD CALL_CORRECTIONPOS
END_METHOD

METHOD CALL_CORRECTIONPROFILE
END_METHOD

METHOD CALL_ENABLEREGISTERCONTROL
END_METHOD

METHOD CALL_ERRORHANDLER
END_METHOD

METHOD CALL_FB
VAR_IN_OUT
	YAXIS : AXIS_REF;
END_VAR
END_METHOD

METHOD CALL_GEARFACTORCORRECTION
END_METHOD

METHOD CALL_GEARING
END_METHOD

METHOD CALL_INPUT
END_METHOD

METHOD CALL_LIMIT
END_METHOD

METHOD CALL_MARKDISTCHANGE
END_METHOD

METHOD CALL_MARKSENSORPOS
END_METHOD

METHOD CALL_MARKSTACK
END_METHOD

METHOD CALL_MARKWINDOW
VAR_IN_OUT
	YAXIS : AXIS_REF;
END_VAR
END_METHOD

METHOD CALL_NOTENABLE
END_METHOD

METHOD CALL_OUTPUT
END_METHOD

METHOD CALL_RESET
END_METHOD

METHOD CALL_RESETOUTPUTS
END_METHOD

METHOD CALL_SETAXISREFMASTERVALUES
END_METHOD

METHOD CALL_TPCONVERTER
END_METHOD

METHOD CALL_VIRTUALACTPOS
END_METHOD

METHOD GET_ACTMARKERRORLIMITED : LREAL
END_METHOD

METHOD GET_ACTUALMARKDIST : LREAL
END_METHOD

METHOD GET_CORRREGPOS : LREAL
END_METHOD

METHOD GET_INTEGRATORREGPOS : LREAL
END_METHOD

METHOD GET_MARKERRORUNLIMITED : LREAL
END_METHOD

METHOD GET_MARKPOSITIONINREGISTER : LREAL
END_METHOD

METHOD GET_MARKRECEIVEUNLIMITED : BOOL
END_METHOD

METHOD GET_MARKRECEIVEDLIMITED : BOOL
END_METHOD

METHOD GET_MARKWINDOWCOMP : BOOL
END_METHOD

METHOD GET_REGISTERINPUTVEL : LREAL
END_METHOD

METHOD GET_SETVELOCITYREGISTER : LREAL
END_METHOD

METHOD GET_LRMARKSTACKLENGTH : LREAL
END_METHOD

METHOD SETTPCOMPFACTOR : LREAL
END_METHOD

METHOD SETTPDELAYCYCLE : LREAL
END_METHOD

(* ---- L_TS2P_MATERIALCOUNTER.pou ---- *)
FUNCTION_BLOCK L_TS2P_MATERIALCOUNTER
VAR_INPUT
	XENABLE : BOOL;
	LRPOSIN : LREAL;
	LRTASKCYCLE : LREAL;
	LRPOSINSLAVE : LREAL;
	LRCYCLELEN : LREAL;
	XLOADSTARTPOS : BOOL;
	XSETMATERIALCOUNTER : BOOL;
	LRSETMATERIALPOS : LREAL;
	XLOADDELTAPOS : BOOL;
	LRSETDELTAPOS : LREAL;
	XSTARTFLYINGSAW : BOOL;
END_VAR
VAR_OUTPUT
	LNMATERIALPOS_E8 : LINT;
	LRMATERIALCOUNTER : LREAL;
	LRDELTAMATERIALPOS : LREAL;
END_VAR
VAR_IN_OUT
	AXIS : AXIS_REF;
END_VAR
VAR
	LNMODULOPOS_E8 : LINT;
	LNMODULOPOSOLD_E8 : LINT;
	LNCYCLELEN_E8 : LINT;
	LNPOSXDIFF : LINT;
	LNMATERIALPOS_E8_OLD : LINT;
	LNDELTAMATERIALPOS : LINT;
	XSETMATERIALCOUNTER_OLD : BOOL;
	XENABLE_OLD : BOOL;
END_VAR
END_FUNCTION_BLOCK

(* ---- L_TS2P_MULTICAMSEQUENCER.pou ---- *)
FUNCTION_BLOCK L_TS2P_MULTICAMSEQUENCER
VAR_INPUT
	XENABLE : BOOL;
	XCAMSEQUENCER : BOOL;
	EMODE : L_TS2P_CamSequenceMode;
	XCAMCHANGEINSTANT : BOOL;
	XLOADCAMTABLE : BOOL;
	WSETCAMTABLE : WORD;
	XENDOFPROFILEIN : BOOL;
	CAMTABLE1 : MC_CAM_REF;
	CAMTABLE2 : MC_CAM_REF;
	CAMTABLE3 : MC_CAM_REF;
	CAMTABLE4 : MC_CAM_REF;
END_VAR
VAR_OUTPUT
	XDONE : BOOL;
	XBUSY : BOOL;
	XERROR : BOOL;
	EERRORID : L_IE1P_Error;
	WACTIVECAMTABLE : WORD;
	CAMTABLEOUT : MC_CAM_REF;
	XCAMTABLEVALID : BOOL;
END_VAR
VAR
	WFMSTATE : WORD := 0;
	XINITSTATE : BOOL;
	XENABLE_OLD : BOOL;
	XLOADCAMTABLE_OLD : BOOL;
	XENDOFPROFILEIN_OLD : BOOL;
	XCAMSEQUENCER_OLD : BOOL;
	XCAMCHANGEINSTANT_OLD : BOOL;
	XCAMSEQUENCERACTIVE : BOOL;
END_VAR
END_FUNCTION_BLOCK

METHOD CALL_ERRORHANDLER
END_METHOD

METHOD CALL_FBMETHODS
END_METHOD

METHOD CALL_OUTPUT
END_METHOD

METHOD CALL_RESETCOMMANDS
END_METHOD

METHOD CALL_RESETOUTPUT
END_METHOD

METHOD CALL_STATEMACHINE
END_METHOD

METHOD CALL_SETCAMTABLEOUT
VAR_INPUT
	WSETCAMTABLE : WORD;
END_VAR
END_METHOD

METHOD CAMREFCHANGED : BOOL
VAR_IN_OUT
	CAMREFNEW : MC_CAM_REF;
	CAMREFOLD : MC_CAM_REF;
END_VAR
END_METHOD

METHOD SET_INIT
END_METHOD

METHOD CALL_S000_CYCLIC
END_METHOD

METHOD CALL_S001_INIT
END_METHOD

METHOD CALL_S002_READY
END_METHOD

METHOD CALL_S151_SEQUENCE_CYCLICCAM1
END_METHOD

METHOD CALL_S152_SEQUENCE_CYCLICCAM3
END_METHOD

METHOD CALL_S153_SEQUENCE_CAM1CYCLICCAM3CAM1
END_METHOD

METHOD CALL_S154_SEQUENCE_CAM1CAM2CYCLICCAM3CAM4CAM1
END_METHOD

(* ---- L_TS2P_OFFSETANDTRIM.pou ---- *)
FUNCTION_BLOCK L_TS2P_OFFSETANDTRIM
VAR_INPUT
	XENABLE : BOOL;
	LRSETOFFSET : LREAL;
	XLOADOFFSET : BOOL;
	XTRIMVELOCITY : BOOL;
	XTRIMPOS : BOOL;
	XTRIMNEG : BOOL;
	XRESETTRIMOFFSET : BOOL;
	EALLOWEDDIRECTION : L_TB2P_AllowedDirection;
	EACTDIRECTION : MC_DIRECTION;
	LRSETTRIMDISTANCE : LREAL;
	LRSETOFFSETTRIMVEL : LREAL := 100.0;
	LRSETOFFSETTRIMACC : LREAL := 1000.0;
	LRSETOFFSETTRIMDEC : LREAL := 1000.0;
	LRSETOFFSETTRIMJERK : LREAL := 100000.0;
	LRCYCMASTERPOS : LREAL;
	LRCYCMASTERVEL : LREAL;
	LRCYCMASTERACC : LREAL;
END_VAR
VAR_OUTPUT
	XBUSY : BOOL;
	XDONE : BOOL;
	XERROR : BOOL;
	EERRORID : WORD;
	LRSETOFFSETOUTTOTAL : LREAL;
	LRSETOFFSETOUT : LREAL;
	LRSETOFFSETOUTTRIM : LREAL;
	LRSETOFFSETOUTTOTALVEL : LREAL;
END_VAR
VAR
	XTRIMPOSOLD : BOOL := FALSE;
	XTRIMNEGOLD : BOOL := FALSE;
	XRESETTRIMOFFSETOLD : BOOL := FALSE;
	LRTRIMPOSITION : LREAL;
	XTRIMPOSEDGE : BOOL;
	XTRIMNEGEDGE : BOOL;
	XABORTPROFILEGENERATORTRIM : BOOL;
	LRTRIMDECDIST : LREAL;
	LRSETOFFSETTRIM_INT : LREAL;
	LRTARGETPOSOLD : LREAL;
	LRSETOFFSETTOTAL : LREAL;
	XPROFILEGENERATORACTIVEOFFSET : BOOL := FALSE;
	LRSETOFFSETOLD : LREAL;
	LRSETOFFSET_INT : LREAL;
	LRSETOFFSETOUTTOTALSAVE : LREAL;
	LRSETOFFSETSAVE : LREAL;
	LRSETPOSOUT_INT : LREAL;
	LRSETVELOUT_INT : LREAL;
	LRSETACCOUT_INT : LREAL;
	LRSETOFFSETTRIMVEL_INT : LREAL;
	LRSETOFFSETTRIMACC_INT : LREAL;
	LRSETOFFSETTRIMDEC_INT : LREAL;
	LRSETOFFSETTRIMJERK_INT : LREAL;
	LRSETOFFSETTRIMVELOLD_INT : LREAL;
	LRSETOFFSETTRIMACCOLD_INT : LREAL;
	LRSETOFFSETTRIMDECOLD_INT : LREAL;
	LRSETOFFSETTRIMJERKOLD_INT : LREAL;
	XMASTERVELDISABLEDDIRECTION : BOOL := FALSE;
	XMASTERVELDISABLEDDIRECTIONOLD : BOOL;
	XEXECUTEPOSITIONING : BOOL;
	XABORTPOSITIONING : BOOL;
	XAUXEXECUTE : BOOL;
	XABORTPOSITIVE : BOOL;
	XINITDONE : BOOL := FALSE;
	LRTASKCYCLETIME : LREAL := 0.001;
	XLOADOFFSET_OLD : BOOL;
	PROFILEGENERATOR : L_MC1P_ProfileGenerator;
	SCPROFILEPARAMETER : L_MC1P_ProfileParameter;
	LRSETOFFSETOUTTOTAL_OLD : LREAL;
END_VAR
END_FUNCTION_BLOCK

METHOD CALL_ADDOFFSETS
END_METHOD

METHOD CALL_AVOIDREVERSING
END_METHOD

METHOD CALL_INITROUTINE
END_METHOD

METHOD CALL_INPUTS
END_METHOD

METHOD CALL_LOADOFFSET
END_METHOD

METHOD CALL_OUTPUT
END_METHOD

METHOD CALL_PROFILEGENERATOR
END_METHOD

METHOD CALL_RESETOUTPUT
END_METHOD

METHOD CALL_TRIMING
END_METHOD

(* ---- L_TS2P_PROCESSCONTROL.pou ---- *)
FUNCTION_BLOCK L_TS2P_PROCESSCONTROL
VAR_INPUT
	XENABLE : BOOL;
	XSYNCFLYINGSAW : BOOL;
	XSYNCININSTANT : BOOL;
	XEXECUTEFIRSTCUT : BOOL;
	XRESUMETARGETPOS : BOOL;
	XRESET : BOOL;
	XTPNOTVALID : BOOL;
	XEXECUTEGAP : BOOL;
	XSETCUTTINGLENGTHINSTANT : BOOL;
	XDONEPROFILE : BOOL;
	LRSLAVEPOSIN : LREAL;
	LRLOWERLIMIT : LREAL;
	LRUPPERLIMIT : LREAL;
	LRSTARTPOS : LREAL;
	LRPOSX1 : LREAL;
	LRVELX1 : LREAL;
	LRACCX1 : LREAL;
	LRTASKCYCLE : LREAL;
END_VAR
VAR_OUTPUT
	XEXECUTEPROFILE : BOOL;
	XAUXEXECUTEPROFILE : BOOL;
	XSYNCPOSOUT : BOOL;
	LRPOSX2 : LREAL;
	LRVELX2 : LREAL;
	LRACCX2 : LREAL;
	XCUTTINGACTIVE : BOOL;
	LRTOLERANCE : LREAL;
	XTARGETOUTSIDELOWERLIMIT : BOOL;
	LRRESTTIMETARGETTOLOWERLIMIT : LREAL;
	LRDISTTOTARGET : LREAL;
END_VAR
VAR
	XEXECUTEPROFILE_INT : BOOL;
	XSYNC_INT : BOOL;
	WSTEPPER : WORD;
	XEXECUTEGAP_OLD : BOOL;
	XRESET_OLD : BOOL;
	XSYNCININSTANT_OLD : BOOL;
	XENABLE_OLD : BOOL;
	LRSTARTTHRESHOLD : LREAL;
	XSETCUTTINGLENGTHINSTANT_OLD : BOOL;
	XRESUMETARGETPOS_OLD : BOOL;
	XEXECUTEFIRSTCUT_OLD : BOOL;
	XMATERIALCONSTANTVEL : BOOL;
	LRMATERIALVEL : LREAL;
	LRMATERIALACC : LREAL;
	XSYNCININSTANT_LOCK : BOOL;
END_VAR
END_FUNCTION_BLOCK

(* ---- L_TS2P_SYNCANDCORRECTIONSTATE.pou ---- *)
FUNCTION_BLOCK L_TS2P_SYNCANDCORRECTIONSTATE EXTENDS L_TB2P_TechModuleBase
VAR_INPUT
	XUSEORIGINAL : BOOL;
	XENABLE : BOOL;
	XENABLEOPERATION : BOOL;
	XRESETERROR : BOOL;
	XQSPAPPLICATION : BOOL;
	XABORT : BOOL;
	XJOGPOS : BOOL;
	XJOGNEG : BOOL;
	XHOMEEXECUTE : BOOL;
	LROVERRIDE : LREAL := 1;
	SCCTRLBASICMOTION : L_TB2P_scCtrlBasicMotion;
	SCPAR : L_TS2P_scPar_SyncAndCorrectionState;
	SCACCESSPOINTS : L_TS2P_scAP_SyncAndCorrectionState;
	MASTERVALUES : L_MC1P_IAXIS_REF_MASTERVALUES;
	XSYNCIN : BOOL;
	XSYNCPOSRESTORE : BOOL;
	LRSETBASEVEL : LREAL;
	LRSETOFFSETPOS : LREAL;
	XTRIMPOS : BOOL;
	XTRIMNEG : BOOL;
	XTRIMRESET : BOOL;
	SCTPRECDATA_MARKSENSOR : L_MC1P_TpReceiveData;
	SCTPRECDATA_TOOLSENSOR : L_MC1P_TpReceiveData;
	XTEACHMARKWINDOW : BOOL;
	XTEACHMARKWINDOWTOOL : BOOL;
	XGEARFACTORCORR : BOOL;
	XGEARFACTORCORRHOLD : BOOL;
END_VAR
VAR_OUTPUT
	XREADYFOROPERATION : BOOL;
	XOPERATIONENABLED : BOOL;
	XREADYFORMOTION : BOOL;
	XERROR : BOOL;
	XWARNING : BOOL;
	EERRORID : L_IE1P_Error;
	XSTOACTIVE : BOOL;
	XQSPACTIVE : BOOL;
	XABORTBUSY : BOOL;
	XABORTDONE : BOOL;
	XJOGGINGBUSY : BOOL;
	XHOMINGBUSY : BOOL;
	XHOMINGDONE : BOOL;
	XISHOMED : BOOL;
	ETMSTATE : L_TB2P_States := L_TB2P_States.DISABLED;
	SCSTATUSBASICMOTION : L_TB2P_scStatusBasicMotion;
	LRACTVEL : LREAL;
	LRSETVELOUT : LREAL;
	LRACTPOS : LREAL;
	LRSETPOSOUT : LREAL;
	LRACTFOLLOWINGERROR : LREAL;
	SCSIGNALFLOW : L_TS2P_scSF_SyncAndCorrectionState;
	XSYNCHRONISED : BOOL;
	XACCDECSYNC : BOOL;
	XOFFSETTRIMACTIVE : BOOL;
	XBASEVELOCITYACTIVE : BOOL;
	LROFFSETTOTAL : LREAL;
	LRSETMARKCORROUT : LREAL;
	XMARKWINDOWTEACHED : BOOL;
	LRGEARFACTORCORR : LREAL;
	LRSETTOOLCORROUT : LREAL;
	XMARKWINDOWTEACHEDTOOL : BOOL;
END_VAR
VAR_IN_OUT
	AXIS : AXIS_REF;
END_VAR
VAR
	XINTERNALCONTROLACTIVE_OLD : BOOL;
	ITFCONNECTORSYNCANDCORRECTION : L_TS2P_IConnectorSyncAndCorrection;
	TM_INT : L_TS2P_TM_SyncAndCorrectionState;
	SCPAR_INT : L_TS2P_scPar_SyncAndCorrectionState;
	SCDATA_INT : L_TS2P_scData_TM_SyncAndCorrectionState;
	SCDATASP_INT : L_TS2P_scData_TM_SyncPosBase;
	XUSEORIGINAL_OLD : BOOL;
	_UICALLMFUNIDXINPUT : UINT := 1;
	_UICALLMFUNIDXOUTPUT : UINT := 1;
	_MCCALL : L_UM1P_MCCall;
	_ASCINPUT : ARRAY [1.._MCCall.c_BufferDepthInput] OF L_TS2P_SyncAndCorrectionStateIn;
	_ASCOUTPUT : ARRAY [1.._MCCall.c_BufferDepthOutput] OF L_TS2P_SyncAndCorrectionStateOut;
	_ASCPARCORE : ARRAY [1.._MCCall.c_BufferDepthInput] OF L_TS2P_scPar_SyncAndCorrectionState;
	_ASCACCESSPOINTSCORE : ARRAY [1.._MCCall.c_BufferDepthInput] OF L_TS2P_scAP_SyncAndCorrectionState;
	_ASCSIGNALFLOWCORE : ARRAY [1.._MCCall.c_BufferDepthOutput] OF L_TS2P_scSF_SyncAndCorrectionState;
	_SCINPUTVISU : L_TS2P_SyncAndCorrectionStateIn;
	_PSCINPUTVISU : POINTER TO L_TS2P_SyncAndCorrectionStateIn := ADR(_scInputVisu);
	_PSCOUTPUTVISU : POINTER TO L_TS2P_SyncAndCorrectionStateOut := ADR(_ascOutput[1]);
	_PSCDATAVISU : POINTER TO L_TS2P_scData_TM_SyncAndCorrectionState := ADR(scData_int);
	_PSCDATASPVISU : POINTER TO L_TS2P_scData_TM_SyncPosBase := ADR(scDataSP_int);
	_PSCPARVISU : POINTER TO L_TS2P_scPar_SyncAndCorrectionState := ADR(scPar_int);
	_PSCAPVISU : POINTER TO L_TS2P_scAP_SyncAndCorrectionState;
	_PSCSFVISU : POINTER TO L_TS2P_scSF_SyncAndCorrectionState;
	ITFBASICMOTIONBASE : L_TB2P.L_TB2P_IBasicMotionBase;
	ITFITECHMODULEINTERNAL : L_TB2P_ITechModuleInternal;
	ITFSYNCANDCORRECTIONEXTENSION : L_TS2P_ISyncAndCorrectionState;
	ITFSYNCPOSEXTENSION : L_TS2P_ISyncPosBase;
	LRJERKDEC : LREAL;
	LRJOGGINGJERKDEC : LREAL;
	REMAININGTIMEOFPROFILE : LREAL;
	REMAININGTIMEOFPROFILEAVAILABLE : BOOL;
END_VAR
END_FUNCTION_BLOCK

METHOD CALL_ABC
VAR_INPUT
	ITFTECHMODULE : L_TB2P.L_TB2P_IBasicMotionBase;
	XQSPAPPLICATION : BOOL;
	XHALT : BOOL;
	XABORT : BOOL;
	XHOMEEXECUTE : BOOL;
	XJOGPOS : BOOL;
	XJOGNEG : BOOL;
	XFINISHPOSITIONING : BOOL;
	XMOVEVELEXECUTE : BOOL;
	XMOVEABSEXECUTE : BOOL;
	XMOVERELEXECUTE : BOOL;
	XENABLEOPERATION : BOOL;
	XRESETERROR : BOOL;
	XENABLEPOSITIVE : BOOL;
	XENABLENEGATIVE : BOOL;
	XDISABLESWLIMIT : BOOL;
	LROVERRIDE : LREAL;
	LROVERRIDEACC : LREAL;
	LROVERRIDEJERK : LREAL;
	XRESETHOMEPOSITION : BOOL;
	XCONTINUOUSUPDATE : BOOL;
	LRPOS_DIST : LREAL;
	LRVEL : LREAL;
	LRACC : LREAL;
	LRDEC : LREAL;
	LRJERK : LREAL;
	EDIRECTION : L_TB2P.MC_DIRECTION;
	SCHOMEEXTTP : L_TB2P.MC_TRIGGER_REF;
	XHOMEABSSWITCH : BOOL;
	XSPECIALABORTBEHAVIOR : BOOL;
	LRABORTDEC : LREAL;
	LRABORTJERK : LREAL;
END_VAR
VAR_OUTPUT
	XERROR : BOOL;
	EERRORID : L_TB2P.L_IE1P_Error;
	XFUNBUSY : BOOL;
	XFUNDONE : BOOL;
	XFUNCOMMANDABORTED : BOOL;
	EFUNSTATEACT : L_TB2P.L_MC1P_ABC_State;
	ECONTROLMODE : L_TB2P.L_MC1P_ControlMode;
	XISHOMED : BOOL;
	XHWLIMITSWITCHNEG : BOOL;
	XHWLIMITSWITCHPOS : BOOL;
	XSWLIMITENABLED : BOOL;
	XSWLIMITSWITCHNEG : BOOL;
	XSWLIMITSWITCHPOS : BOOL;
	EAXISTYPE : L_TB2P.L_MC1P_DriveType;
	EAXISSTATE : L_TB2P.L_MC1P_AXIS_STATE;
	XSTOACTIVE : BOOL;
	XREADYFOROPERATION : BOOL;
	XOPERATIONENABLED : BOOL;
	XREADYFORMOTION : BOOL;
	XAXISWARNING : BOOL;
	XAXISERROR : BOOL;
	EAXISERRORID : L_TB2P.L_IE1P_Error;
	XDRIVEWARNING : BOOL;
	XDRIVEERROR : BOOL;
	DWDRIVEERRORID : DWORD;
	LRACTPOS : LREAL;
	LRACTVEL : LREAL;
	LRSETPOSOUT : LREAL;
	LRSETVELOUT : LREAL;
	LRACTFOLLOWINGERROR : LREAL;
	XINPOSITION : BOOL;
	XSTANDSTILLSETVELOCITY : BOOL;
	XSTANDSTILLACTVELOCITY : BOOL;
	XCONSTANTVELOCITY : BOOL;
	XACCELERATING : BOOL;
	XDECELERATING : BOOL;
	XDIRECTIONPOSITIVE : BOOL;
	XDIRECTIONNEGATIVE : BOOL;
	XAXISAVAILABLE : BOOL;
END_VAR
VAR_IN_OUT
	AXIS : AXIS_REF;
END_VAR
END_METHOD

METHOD GET_PAP : POINTER TO L_TB2P_scAP_TM_MotionControl
END_METHOD

METHOD GET_PDATA : POINTER TO L_TS2P_scData_TM_SyncAndCorrectionState
END_METHOD

METHOD GET_PDATASP : POINTER TO L_TS2P_scData_TM_SyncPosBase
END_METHOD

METHOD GET_PPAR : POINTER TO L_TB2P.L_TB2P_scPar_TM_MotionControl
END_METHOD

METHOD GET_PSF : POINTER TO L_TB2P_scSF_TM_MotionControl
END_METHOD

METHOD ADDOFFSET
VAR_INPUT
	ITFTECHMODULE : L_TS2P_ISyncPosBase;
	LRSETPOS : LREAL;
	LRSETVEL : LREAL;
	LRSETOFFSET : LREAL;
	LRSETOFFSETVEL : LREAL;
	ETRAVERSINGRANGE : L_MC1P.L_MC1P_TraversingRange;
	LRCYCLELENGTH : LREAL;
END_VAR
VAR_OUTPUT
	XERROR : BOOL;
	EERRORID : L_IE1P.L_IE1P_Error;
	LRSETPOSOUT : LREAL;
	LRSETVELOUT : LREAL;
END_VAR
END_METHOD

METHOD CLUTCH
VAR_INPUT
	ITFTECHMODULE : L_TS2P_ISyncPosBase;
	XENABLE : BOOL;
	XSYNCIN : BOOL;
	LRSETBASEVELOCITY : LREAL;
	ESYNCMODE : L_TB2P_SyncMode;
	EALLOWEDDIRECTION : L_TB2P_AllowedDirection;
	LRSYNCVEL : LREAL;
	LRSYNCACC : LREAL;
	LRSYNCDEC : LREAL;
	LRSYNCJERK : LREAL;
	LRSYNCINDIST : LREAL;
	LRSYNCOUTDIST : LREAL;
	LRSYNCOUTPOS : LREAL;
	XLOADCLUTCHOFFSET : BOOL;
	LRLOADCLUTCHOFFSET : LREAL;
	LRCYCLICMASTERPOS : LREAL;
	LRCYCLICMASTERVEL : LREAL;
	ETRAVERSINGRANGEMASTER : L_MC1P_TraversingRange;
	LRCYCLELENGTHMASTER : LREAL;
	LRCYCLICAXISPOS : LREAL;
	LRCYCLICAXISVEL : LREAL;
	LRCYCLICAXISACC : LREAL;
	ETRAVERSINGRANGEAXIS : L_MC1P_TraversingRange;
	LRCYCLELENGTHAXIS : LREAL;
END_VAR
VAR_OUTPUT
	XERROR : BOOL;
	EERRORID : L_IE1P.L_IE1P_Error;
	XBUSY : BOOL;
	XDONE : BOOL;
	XSYNCHRONISED : BOOL;
	XACCDECSYNC : BOOL;
	XINBASEVELOCITY : BOOL;
	LRSETPOSOUT : LREAL;
	LRSETVELOUT : LREAL;
	LRSETACCOUT : LREAL;
	LRCLUTCHOFFSETOUT : LREAL;
END_VAR
END_METHOD

METHOD GEARBOX
VAR_INPUT
	ITFTECHMODULE : L_TS2P_ISyncPosBase;
	XENABLE : BOOL;
	LRSETPOSX : LREAL;
	LRSETVELX : LREAL;
	DWNUMERATOR : DWORD;
	DWDENOMINATOR : DWORD;
	LRCYCLELENGTHX : LREAL;
	LRCYCLELENGTHY : LREAL;
	ETRAVERSINGRANGEX : L_MC1P.L_MC1P_TraversingRange;
	ETRAVERSINGRANGEY : L_MC1P.L_MC1P_TraversingRange;
	XLOADGEARBOXPOS : BOOL;
	LRLOADGEARBOXPOS : LREAL;
END_VAR
VAR_OUTPUT
	XERROR : BOOL;
	EERRORID : L_IE1P.L_IE1P_Error;
	LRSETPOSOUT : LREAL;
	LRSETVELOUT : LREAL;
END_VAR
END_METHOD

METHOD OFFSETANDTRIM
VAR_INPUT
	ITFTECHMODULE : L_TS2P_ISyncPosBase;
	XENABLE : BOOL;
	LRSETOFFSET : LREAL;
	XTRIMPOS : BOOL;
	XTRIMNEG : BOOL;
	LRSETTRIMDISTANCE : LREAL;
	ETRIMMODE : L_TS2P_TrimMode;
	XLOADOFFSET : BOOL;
	XRESETTRIMOFFSET : BOOL;
	LRSETVEL : LREAL;
	LRSETACC : LREAL;
	LRSETDEC : LREAL;
	LRSETJERK : LREAL;
	WACTDIRECTION : WORD;
	EALLOWEDDIRECTION : L_TB2P.L_TB2P_AllowedDirection;
	LRCYCMASTERPOS : LREAL;
	LRCYCMASTERVEL : LREAL;
	LRCYCMASTERACC : LREAL;
END_VAR
VAR_OUTPUT
	XERROR : BOOL;
	EERRORID : L_IE1P.L_IE1P_Error;
	XBUSY : BOOL;
	XDONE : BOOL;
	LRSETOFFSETOUTTOTAL : LREAL;
	LRSETOFFSETOUTTOTALVEL : LREAL;
	LRSETOFFSETOUT : LREAL;
	LRSETOFFSETOUTTRIM : LREAL;
END_VAR
END_METHOD

METHOD REQUESTINTERFACE : BOOL
VAR_INPUT
	ID : DINT;
	PITFUNKNOWN : POINTER TO L_UBUP.L_UBUP_IUnknown;
END_VAR
END_METHOD

METHOD CALLFUNCTION
VAR_INPUT
	UIINPUTDATAIDX : UINT;
	UIOUTPUTDATAIDX : UINT;
END_VAR
END_METHOD

METHOD COPYINPUTS : BOOL
VAR_INPUT
	IDX : WORD;
END_VAR
END_METHOD

METHOD COPYOUTPUTS : BOOL
VAR_INPUT
	IDX : WORD;
END_VAR
END_METHOD

METHOD FUNCTIONWASCALLEDTWICE : BOOL
VAR_INPUT
	IDX : WORD;
END_VAR
END_METHOD

METHOD HANDLESTANDARDCALL : BOOL
END_METHOD

METHOD SYNCOUTPUTS
VAR_INPUT
	UICOPYOUTPUTFROMIDX : UINT;
	UICOPYOUTPUTTOIDX : UINT;
END_VAR
END_METHOD

METHOD FB_INIT : BOOL
VAR_INPUT
	BINITRETAINS : BOOL;
	BINCOPYCODE : BOOL;
END_VAR
END_METHOD

METHOD CALL_INTERNALCTRL
END_METHOD

(* ---- L_TS2P_SYNCDRIVEPOS.pou ---- *)
FUNCTION_BLOCK L_TS2P_SYNCDRIVEPOS
VAR_INPUT
	MASTERAXIS : POINTER TO L_MC1P_IAXIS_REF_MASTERVALUES;
	XENABLE : BOOL;
	DWNUMERATOR : DWORD := 1;
	DWDENOMINATOR : DWORD := 1;
	XSYNCIN : BOOL;
	XSYNCOUTINSTANT : BOOL;
	XSYNCINSTANT : BOOL;
	XCLUTCHRELATIVE : BOOL;
	XSYNCPOSRESTORE : BOOL;
	LRSLAVESYNCOUTPOS : LREAL;
	LRSLAVESYNCINDIST : LREAL := 90;
	LRSLAVESYNCOUTDIST : LREAL := 90;
	LRSYNCOUTINSTANTDEC : LREAL := 10000;
	EALLOWEDDIRECTION : L_TB2P_AllowedDirection := L_TB2P_AllowedDirection.both;
	ESYNCMODE : L_TB2P_SyncMode := L_TB2P_SyncMode.ProfGenAbsolute;
	LRSYNCVEL : LREAL := 100;
	LRSYNCACC : LREAL := 1000.0;
	LRSYNCDEC : LREAL := 1000.0;
	LRSYNCJERK : LREAL := 10000000000.0;
	LRSETBASEVELOCITY : LREAL := 0;
	XLOADCLUTCHOFFSET : BOOL := FALSE;
	LRLOADCLUTCHOFFSET : LREAL := 0;
	XTRIMVELOCITYX : BOOL;
	XTRIMVELOCITYY : BOOL;
	LRSETTRIMDISTANCEX : LREAL := 1;
	LRSETTRIMDISTANCEY : LREAL := 1;
	XTRIMPOSX : BOOL;
	XTRIMNEGX : BOOL;
	XTRIMPOSY : BOOL;
	XTRIMNEGY : BOOL;
	XRESETTRIMX : BOOL;
	XRESETTRIMY : BOOL;
	LRSETOFFSETX : LREAL := 0;
	LRSETOFFSETTRIMVELX : LREAL := 10.0;
	LRSETOFFSETTRIMACCX : LREAL := 100.0;
	LRSETOFFSETTRIMDECX : LREAL := 100.0;
	LRSETOFFSETTRIMJERKX : LREAL := 10000.0;
	XLOADOFFSETX : BOOL;
	LRSETOFFSETY : LREAL := 0;
	LRSETOFFSETTRIMVELY : LREAL := 10.0;
	LRSETOFFSETTRIMACCY : LREAL := 100.0;
	LRSETOFFSETTRIMDECY : LREAL := 100.0;
	LRSETOFFSETTRIMJERKY : LREAL := 10000.0;
	XLOADOFFSETY : BOOL;
	XLOADSTARTSLAVEPOS : BOOL := FALSE;
	LRSTARTSLAVEPOS : LREAL;
	XLOADGEARBOXPOS : BOOL;
	LRLOADGEARBOXPOS : LREAL;
	XOPERATIONENABLED : BOOL;
END_VAR
VAR_OUTPUT
	XERROR : BOOL;
	XWARNING : BOOL;
	EERRORID : L_IE1P_Error;
	XBUSY : BOOL;
	LRSETSLAVEPOSOUT : LREAL;
	LRSETSLAVEVELOUT : LREAL;
	LRSETSLAVEACCOUT : LREAL;
	LRSETGEARBOXPOSOUT : LREAL;
	XSYNCOUTDONE : BOOL;
	XSYNCHRONISED : BOOL;
	XACCDECSYNC : BOOL;
	XOFFSETTRIMBUSY : BOOL;
	LROFFSETOUTTOTALVELX : LREAL;
	LROFFSETOUTTOTALVELY : LREAL;
	LROFFSETOUTTRIMX : LREAL;
	LROFFSETOUTTRIMY : LREAL;
	LROFFSETOUTX : LREAL;
	LROFFSETOUTY : LREAL;
	LROFFSETOUTTOTALX : LREAL;
	LROFFSETOUTTOTALY : LREAL;
	LRSETCLUTCHPOS : LREAL;
	LRSETCLUTCHVEL : LREAL;
	LRSETCLUTCHACC : LREAL;
	XBASEVELSYNCHRONISED : BOOL;
	XACCDECBASEVEL : BOOL;
	LROFFSETSYNCPOS : LREAL;
END_VAR
VAR_IN_OUT
	SLAVEAXIS : AXIS_REF;
END_VAR
VAR
	FB_GEARBOXPOSITION : L_MB1P_GearboxPositionInput;
	FB_CLUTCHEXTENDEDBASE : L_TB2P_ClutchExtendedBase;
	FB_AXISCONVERTER : L_MC2P.L_MC2P_AxisConverterBase;
	FB_OFFSETANDTRIMX : L_TS2P_OffsetAndTrim;
	FB_ADDOFFSETCYCLICX : L_MC1P_AddOffsetCyclic;
	FB_OFFSETANDTRIMY : L_TS2P_OffsetAndTrim;
	FB_ADDOFFSETCYCLICY : L_MC1P_AddOffsetCyclic;
	FB_SYNCPOSRESTOREOFFSET : L_TS2P_OffsetAndTrim;
	FB_DIRECTION : L_MC1P_GetDirection;
	LRSETOFFSETMASTER_INT : LREAL;
	LRTRIMDIST_INT : LREAL;
	XTRIMPOS_OLD : BOOL;
	XTRIMNEG_OLD : BOOL;
	XTRIMVEL : BOOL;
	LRTRIMOFFSETDIST : LREAL;
	LRLOADOFFSETMASTER_INT : LREAL := 0;
	LRLOADGEARBOXPOS_INT : LREAL;
	LRSETGEARBOXPOSOUT_INT : LREAL;
	XSETDISABLECLUTCH_INT : BOOL;
	LRLOADTRIMOFFSET_INT : LREAL := 0;
	LRSYNCOUTINSTANTDEC_INT : LREAL := 100000;
	LRSETINTEGRATETRIMVELPOSOUT_INT : LREAL;
	XSYNCPOS_OLD : BOOL;
	XRESETTRIM_OLD : BOOL;
	LRLOADOFFSET_INT : LREAL := 0;
	XSYNCINSTANT_OLD : BOOL;
	XENABLEGEARBOX : BOOL;
	LRSYNCOFFSET : LREAL;
	LRSCALING_INT : LREAL := 1;
	LRGEARBOXSTARTPOSOUT_INT : LREAL;
	DWDENOMINATOR_INT : DWORD := 1;
	XENABLE_OLD : BOOL;
	WAXESMODE : WORD;
	WAXESMODEOLD : WORD;
	LRADDOFFSETPOSOUTY_OLD : LREAL;
	LRADDOFFSETVELOUTY : LREAL;
	LRSETGEARBOXPOSOUTOLD_INT : LREAL;
	LRSETGEARBOXPOSOUTVEL_INT : LREAL;
	LRGETGEARBOXVELIN : LREAL;
	LRGETGEARBOXPOSOUT : LREAL;
	LRGETGEARBOXPOSIN : LREAL;
	LRTASKCYCLE : LREAL;
	XINIT : BOOL := TRUE;
	XCLUTCHDONE_OLD : BOOL;
	XENABLEOLD : BOOL;
	LRSETOFFSETOUTTOTALVELOLD : LREAL;
	SET_AP_LRMASTERVELSTANDSTILLDEADBAND : LREAL;
END_VAR
END_FUNCTION_BLOCK

METHOD CALL_AXESMODE
END_METHOD

METHOD CALL_CALCGEARBOXOUTVELACC
VAR_IN_OUT
	SLAVEAXIS : AXIS_REF;
END_VAR
END_METHOD

METHOD CALL_ERRORHANDLER
END_METHOD

METHOD CALL_FBMETHODS
END_METHOD

METHOD CALL_FBMETHODS_FMDISABLE
END_METHOD

METHOD CALL_FB_ADDOFFSETCYCLICX
END_METHOD

METHOD CALL_FB_ADDOFFSETCYCLICX_INPUT
END_METHOD

METHOD CALL_FB_ADDOFFSETCYCLICY
END_METHOD

METHOD CALL_FB_ADDOFFSETCYCLICY_INPUT
END_METHOD

METHOD CALL_FB_AXISCONVERTER
END_METHOD

METHOD CALL_FB_AXISCONVERTER_INPUT
END_METHOD

METHOD CALL_FB_CLUTCHEXTENDEDBASE
END_METHOD

METHOD CALL_FB_CLUTCHEXTENDEDBASE_INPUT
END_METHOD

METHOD CALL_FB_CLUTCHEXTENDEDBASE_INPUTMASTER
END_METHOD

METHOD CALL_FB_CLUTCHEXTENDEDBASE_INPUTSLAVE
VAR_IN_OUT
	SLAVEAXIS : AXIS_REF;
END_VAR
END_METHOD

METHOD CALL_FB_GEARBOXPOSITION
END_METHOD

METHOD CALL_FB_GEARBOXPOSITION_INPUT
END_METHOD

METHOD CALL_FB_GEARBOXPOSITION_LOADGEARBOXPOS
END_METHOD

METHOD CALL_FB_SYNCPOSRESTOREOFFSET
END_METHOD

METHOD CALL_FB_SYNCPOSRESTOREOFFSET_INPUT
VAR_IN_OUT
	SLAVEAXIS : AXIS_REF;
END_VAR
END_METHOD

METHOD CALL_LOADSLAVESTARTPOS
END_METHOD

METHOD CALL_OFFSETANDTRIMX
END_METHOD

METHOD CALL_OFFSETANDTRIMX_INPUT
END_METHOD

METHOD CALL_OFFSETANDTRIMY
END_METHOD

METHOD CALL_OFFSETANDTRIMY_INPUT
END_METHOD

METHOD CALL_OUTPUT
END_METHOD

METHOD CALL_OUTPUT_CLUTCHSTATE
END_METHOD

METHOD CALL_OUTPUT_OFFSET
END_METHOD

METHOD CALL_RESETCOMMANDS
END_METHOD

METHOD CALL_INIT
VAR_IN_OUT
	SLAVEAXIS : AXIS_REF;
END_VAR
END_METHOD

METHOD GET_DIRECTION
END_METHOD

METHOD GET_GETGEARBOXPOSIN : LREAL
END_METHOD

METHOD GET_GETGEARBOXPOSOUT : LREAL
END_METHOD

METHOD GET_GETGEARBOXVELIN : LREAL
END_METHOD

METHOD GET_GETGEARBOXVELOUT : LREAL
END_METHOD

METHOD GET_LRCLUTCHPOSIN : LREAL
END_METHOD

METHOD GET_LROFFSETADDOFFSETCYCLIC : LREAL
END_METHOD

METHOD SETDISABLECLUTCH : BOOL
VAR_INPUT
	XSETDISABLECLUTCH : BOOL;
END_VAR
END_METHOD

(* ---- L_TS2P_SYNCDRIVEVEL.pou ---- *)
FUNCTION_BLOCK L_TS2P_SYNCDRIVEVEL
VAR_INPUT
	MASTERAXIS : POINTER TO L_MC1P_IAXIS_REF_MASTERVALUES;
	XENABLE : BOOL;
	LRCOUPLINGX : LREAL := 1.0;
	LRCOUPLINGY : LREAL := 1.0;
	XINVERTGEARFACTOR : BOOL;
	XDISABLETOLERANCEINVERTGEARFACTOR : BOOL;
	LRTOLERANCEINVERTGEARFACTOR : LREAL := 0;
	XSYNCIN : BOOL;
	XSYNCOUTINSTANT : BOOL;
	LRSYNCACC : LREAL := 10.0;
	LRSYNCDEC : LREAL := 10.0;
	LRSYNCOUTINSTANTDEC : LREAL := 100.0;
	LRSYNCJERK : LREAL := 1.0;
	XAVOIDVELGAPS : BOOL;
	LRSETOFFSETVEL : LREAL;
	DWMODE : DWORD := 1;
	XTRIMVELOCITYX : BOOL;
	XTRIMVELOCITYY : BOOL;
	LRSETTRIMDISTANCEX : LREAL := 1;
	LRSETTRIMDISTANCEY : LREAL := 1;
	XTRIMPOSX : BOOL;
	XTRIMNEGX : BOOL;
	XTRIMPOSY : BOOL;
	XTRIMNEGY : BOOL;
	XRESETTRIMX : BOOL;
	XRESETTRIMY : BOOL;
	XSYNCVELRESET : BOOL;
	LRSETOFFSETX : LREAL := 0;
	LRSETOFFSETTRIMVELX : LREAL := 10.0;
	LRSETOFFSETTRIMACCX : LREAL := 100.0;
	LRSETOFFSETTRIMDECX : LREAL := 100.0;
	LRSETOFFSETTRIMJERKX : LREAL := 10000.0;
	XLOADOFFSETX : BOOL;
	LRSETOFFSETY : LREAL := 0;
	LRSETOFFSETTRIMVELY : LREAL := 10.0;
	LRSETOFFSETTRIMACCY : LREAL := 100.0;
	LRSETOFFSETTRIMDECY : LREAL := 100.0;
	LRSETOFFSETTRIMJERKY : LREAL := 10000.0;
	XLOADOFFSETY : BOOL;
	EALLOWEDDIRECTION : L_TB2P_AllowedDirection;
	XLOADOFFSET : BOOL;
	XLOADGROUNDVEL : BOOL;
	LRSETGROUNDVEL : LREAL;
	LRGROUNDVELACC : LREAL := 10.0;
	LRGROUNDVELDEC : LREAL := 10.0;
	LRGROUNDVELJERK : LREAL := 1.0;
END_VAR
VAR_OUTPUT
	XERROR : BOOL;
	XWARNING : BOOL;
	EERRORID : L_IE1P_Error;
	XBUSY : BOOL;
	LRSETSLAVEVELOUT : LREAL;
	LRSETSLAVEACCOUT : LREAL;
	XSYNCOUTDONE : BOOL;
	XSYNCHRONISED : BOOL;
	XACCDECSYNC : BOOL;
	XOFFSETTRIMBUSY : BOOL;
	LRPOSOFFSETOUTTRIMX : LREAL;
	LRPOSOFFSETOUTTRIMY : LREAL;
	LRPOSOFFSETOUTX : LREAL;
	LRPOSOFFSETOUTY : LREAL;
	LRPOSOFFSETOUTVELX : LREAL;
	LRVELOFFSET : LREAL;
	LROFFSETOUTTOTALX : LREAL;
	LROFFSETOUTTOTALY : LREAL;
	LROFFSETOUTTOTALVELX : LREAL;
	LROFFSETOUTTOTALVELY : LREAL;
	XBASEVELSYNCHRONISED : BOOL;
	XACCDECBASEVEL : BOOL;
	XBASEVELSYNCOUTDONE : BOOL;
	XINVERTGEARFACTORACTIVE : BOOL;
END_VAR
VAR_IN_OUT
	SLAVEAXIS : AXIS_REF;
END_VAR
VAR
	XENABLE_OLD : BOOL;
	ESTATE : L_TF1P_States := L_TF1P_States.INIT;
	ESTATE_OLD : L_TF1P_States := L_TF1P_States.INIT;
	XSTATEENTRY : BOOL;
	FB_CONVAXISV : L_MC2P_ConvAxisV;
	FB_INVERTGEARFACTOR : L_TS2P_InvertGearfactor;
	XACCDECSYNC_OLD : BOOL;
	XSYNCVEL_OLD : BOOL;
	XOPEN_OLD : BOOL;
	LRSETVELTRIM : LREAL;
	XSETDISABLECLUTCH_INT : BOOL;
	SETPOSITIONFORSYNCOLD : LREAL := 0;
	XINITFB_CLUTCHV : BOOL;
	FB_CLUTCHV : L_MC2P_ClutchVelocity;
	XINVERTGEARFACTORACTIVE_OLD : BOOL;
	LRSETGROUNDVEL_INT : LREAL;
	FB_OFFSETANDTRIMX : L_TS2P_OffsetAndTrim;
	FB_VELOCITYOFFSET : L_MC1P_RampGenerator;
	FB_OFFSETANDTRIMY : L_TS2P_OffsetAndTrim;
	FB_RAMPGENGROUNDVEL : L_MC1P_RampGenerator;
	FB_DIRECTION : L_MC1P_GetDirection;
END_VAR
END_FUNCTION_BLOCK

METHOD CALL_ERRORHANDLER
END_METHOD

METHOD CALL_FBMETHODS
END_METHOD

METHOD CALL_FBMETHODS_FMDISABLE
END_METHOD

METHOD CALL_FB_CLUTCHV
END_METHOD

METHOD CALL_FB_CLUTCHV_INPUT
END_METHOD

METHOD CALL_FB_CLUTCHV_PAR
END_METHOD

METHOD CALL_FB_CONVAXISV
END_METHOD

METHOD CALL_FB_CONVAXISV_INPUT
END_METHOD

METHOD CALL_FB_INVERTGEARFACTOR
END_METHOD

METHOD CALL_FB_INVERTGEARFACTOR_INPUT
END_METHOD

METHOD CALL_FB_RAMPGENGROUNDVEL
END_METHOD

METHOD CALL_FB_RAMPGENGROUNDVEL_INPUT
END_METHOD

METHOD CALL_FB_VELOCITYOFFSET
END_METHOD

METHOD CALL_FB_VELOCITYOFFSET_INPUT
END_METHOD

METHOD CALL_OFFSETANDTRIMX
END_METHOD

METHOD CALL_OFFSETANDTRIMX_INPUT
END_METHOD

METHOD CALL_OFFSETANDTRIMY
END_METHOD

METHOD CALL_OFFSETANDTRIMY_INPUT
END_METHOD

METHOD CALL_OUTPUT
END_METHOD

METHOD CALL_OUTPUT_SETSLAVEOUT
END_METHOD

METHOD CALL_RESETCOMMANDS
END_METHOD

METHOD CALL_RESETFM
END_METHOD

METHOD CALL_RESETOUTPUT
END_METHOD

METHOD CALL_STATEMASHINE
END_METHOD

METHOD GET_DIRECTION
END_METHOD

METHOD GET_CLUTCHVELOUT : LREAL
END_METHOD

METHOD GET_GETGEARBOXVELIN : LREAL
END_METHOD

METHOD GET_GETGEARBOXVELOUT : LREAL
END_METHOD

METHOD SETDISABLECLUTCH : BOOL
VAR_INPUT
	XSETDISABLECLUTCH : BOOL;
END_VAR
END_METHOD

METHOD CALL_S000_CYCLIC
END_METHOD

METHOD CALL_S001_INIT
END_METHOD

METHOD CALL_S010_READY
END_METHOD

METHOD CALL_S998_ERROR
END_METHOD

(* ---- L_TS2P_SYNCPOSBASE.pou ---- *)
FUNCTION_BLOCK L_TS2P_SYNCPOSBASE EXTENDS L_TB2P_TechModuleBase
VAR_INPUT
	XUSEORIGINAL : BOOL;
	XENABLE : BOOL;
	XENABLEOPERATION : BOOL;
	XRESETERROR : BOOL;
	XQSPAPPLICATION : BOOL;
	XABORT : BOOL;
	XJOGPOS : BOOL;
	XJOGNEG : BOOL;
	XHOMEEXECUTE : BOOL;
	LROVERRIDE : LREAL := 1;
	SCCTRLBASICMOTION : L_TB2P_scCtrlBasicMotion;
	SCPAR : L_TS2P_scPar_SyncPosBase;
	SCACCESSPOINTS : L_TS2P_scAP_SyncPosBase;
	MASTERVALUES : L_MC1P_IAXIS_REF_MASTERVALUES;
	XSYNCIN : BOOL;
	XSYNCPOSRESTORE : BOOL;
	LRSETBASEVEL : LREAL;
	LRSETOFFSETPOS : LREAL;
	XTRIMPOS : BOOL;
	XTRIMNEG : BOOL;
	XTRIMRESET : BOOL;
END_VAR
VAR_OUTPUT
	XREADYFOROPERATION : BOOL;
	XOPERATIONENABLED : BOOL;
	XREADYFORMOTION : BOOL;
	XERROR : BOOL;
	XWARNING : BOOL;
	EERRORID : L_IE1P_Error;
	XSTOACTIVE : BOOL;
	XQSPACTIVE : BOOL;
	XABORTBUSY : BOOL;
	XABORTDONE : BOOL;
	XJOGGINGBUSY : BOOL;
	XHOMINGBUSY : BOOL;
	XHOMINGDONE : BOOL;
	XISHOMED : BOOL;
	ETMSTATE : L_TB2P_States;
	SCSTATUSBASICMOTION : L_TB2P_scStatusBasicMotion;
	LRACTVEL : LREAL;
	LRSETVELOUT : LREAL;
	LRACTPOS : LREAL;
	LRSETPOSOUT : LREAL;
	LRACTFOLLOWINGERROR : LREAL;
	SCSIGNALFLOW : L_TS2P_scSF_SyncPosBase;
	XSYNCHRONISED : BOOL;
	XACCDECSYNC : BOOL;
	XOFFSETTRIMACTIVE : BOOL;
	XBASEVELOCITYACTIVE : BOOL;
	LROFFSETTOTAL : LREAL;
END_VAR
VAR_IN_OUT
	AXIS : AXIS_REF;
END_VAR
VAR
	XINTERNALCONTROLACTIVE_OLD : BOOL;
	ITFCONNECTORSYNCPOS : L_TS2P_IConnectorSyncPos;
	_XCONNECTORVALID : BOOL;
	TM_INT : L_TS2P_TM_SyncPosBase;
	SCPAR_INT : L_TS2P_scPar_SyncPosBase;
	SCDATA_INT : L_TS2P_scData_TM_SyncPosBase;
	XUSEORIGINAL_OLD : BOOL;
	_UICALLMFUNIDXINPUT : UINT := 1;
	_UICALLMFUNIDXOUTPUT : UINT := 1;
	_MCCALL : L_UM1P_MCCall := STRUCT(itfMCCall := THIS^);
	_ASCINPUT : ARRAY [1.._MCCall.c_BufferDepthInput] OF L_TS2P_SyncPosBaseIn;
	_ASCOUTPUT : ARRAY [1.._MCCall.c_BufferDepthOutput] OF L_TS2P_SyncPosBaseOut;
	_ASCPARCORE : ARRAY [1.._MCCall.c_BufferDepthInput] OF L_TS2P_scPar_SyncPosBase;
	_ASCACCESSPOINTSCORE : ARRAY [1.._MCCall.c_BufferDepthInput] OF L_TS2P_scAP_SyncPosBase;
	_ASCSIGNALFLOWCORE : ARRAY [1.._MCCall.c_BufferDepthOutput] OF L_TS2P_scSF_SyncPosBase;
	_SCINPUTVISU : L_TS2P_SyncPosBaseIn;
	_PSCINPUTVISU : POINTER TO L_TS2P_SyncPosBaseIn := ADR(_scInputVisu);
	_PSCOUTPUTVISU : POINTER TO L_TS2P_SyncPosBaseOut := ADR(_ascOutput[1]);
	_PSCDATAVISU : POINTER TO L_TS2P_scData_TM_SyncPosBase := ADR(scData_int);
	_PSCPARVISU : POINTER TO L_TS2P_scPar_SyncPosBase := ADR(scPar_int);
	_PSCAPVISU : POINTER TO L_TS2P_scAP_SyncPosBase;
	_PSCSFVISU : POINTER TO L_TS2P_scSF_SyncPosBase;
	ITFBASICMOTIONBASE : L_TB2P.L_TB2P_IBasicMotionBase;
	ITFITECHMODULEINTERNAL : L_TB2P_ITechModuleInternal;
	ITFSYNCPOSEXTENSION : L_TS2P_ISyncPosBase;
	LRJERKDEC : LREAL;
	LRJOGGINGJERKDEC : LREAL;
	REMAININGTIMEOFPROFILE : LREAL;
	REMAININGTIMEOFPROFILEAVAILABLE : BOOL;
END_VAR
END_FUNCTION_BLOCK

METHOD CALL_ABC
VAR_INPUT
	ITFTECHMODULE : L_TB2P.L_TB2P_IBasicMotionBase;
	XQSPAPPLICATION : BOOL;
	XHALT : BOOL;
	XABORT : BOOL;
	XHOMEEXECUTE : BOOL;
	XJOGPOS : BOOL;
	XJOGNEG : BOOL;
	XFINISHPOSITIONING : BOOL;
	XMOVEVELEXECUTE : BOOL;
	XMOVEABSEXECUTE : BOOL;
	XMOVERELEXECUTE : BOOL;
	XENABLEOPERATION : BOOL;
	XRESETERROR : BOOL;
	XENABLEPOSITIVE : BOOL;
	XENABLENEGATIVE : BOOL;
	XDISABLESWLIMIT : BOOL;
	LROVERRIDE : LREAL;
	LROVERRIDEACC : LREAL;
	LROVERRIDEJERK : LREAL;
	XRESETHOMEPOSITION : BOOL;
	XCONTINUOUSUPDATE : BOOL;
	LRPOS_DIST : LREAL;
	LRVEL : LREAL;
	LRACC : LREAL;
	LRDEC : LREAL;
	LRJERK : LREAL;
	EDIRECTION : L_TB2P.MC_DIRECTION;
	SCHOMEEXTTP : L_TB2P.MC_TRIGGER_REF;
	XHOMEABSSWITCH : BOOL;
	XSPECIALABORTBEHAVIOR : BOOL;
	LRABORTDEC : LREAL;
	LRABORTJERK : LREAL;
END_VAR
VAR_OUTPUT
	XERROR : BOOL;
	EERRORID : L_TB2P.L_IE1P_Error;
	XFUNBUSY : BOOL;
	XFUNDONE : BOOL;
	XFUNCOMMANDABORTED : BOOL;
	EFUNSTATEACT : L_TB2P.L_MC1P_ABC_State;
	ECONTROLMODE : L_TB2P.L_MC1P_ControlMode;
	XISHOMED : BOOL;
	XHWLIMITSWITCHNEG : BOOL;
	XHWLIMITSWITCHPOS : BOOL;
	XSWLIMITENABLED : BOOL;
	XSWLIMITSWITCHNEG : BOOL;
	XSWLIMITSWITCHPOS : BOOL;
	EAXISTYPE : L_TB2P.L_MC1P_DriveType;
	EAXISSTATE : L_TB2P.L_MC1P_AXIS_STATE;
	XSTOACTIVE : BOOL;
	XREADYFOROPERATION : BOOL;
	XOPERATIONENABLED : BOOL;
	XREADYFORMOTION : BOOL;
	XAXISWARNING : BOOL;
	XAXISERROR : BOOL;
	EAXISERRORID : L_TB2P.L_IE1P_Error;
	XDRIVEWARNING : BOOL;
	XDRIVEERROR : BOOL;
	DWDRIVEERRORID : DWORD;
	LRACTPOS : LREAL;
	LRACTVEL : LREAL;
	LRSETPOSOUT : LREAL;
	LRSETVELOUT : LREAL;
	LRACTFOLLOWINGERROR : LREAL;
	XINPOSITION : BOOL;
	XSTANDSTILLSETVELOCITY : BOOL;
	XSTANDSTILLACTVELOCITY : BOOL;
	XCONSTANTVELOCITY : BOOL;
	XACCELERATING : BOOL;
	XDECELERATING : BOOL;
	XDIRECTIONPOSITIVE : BOOL;
	XDIRECTIONNEGATIVE : BOOL;
	XAXISAVAILABLE : BOOL;
END_VAR
VAR_IN_OUT
	AXIS : AXIS_REF;
END_VAR
END_METHOD

METHOD GET_PAP : POINTER TO L_TB2P_scAP_TM_MotionControl
END_METHOD

METHOD GET_PDATA : POINTER TO L_TS2P_scData_TM_SyncPosBase
END_METHOD

METHOD GET_PPAR : POINTER TO L_TB2P.L_TB2P_scPar_TM_MotionControl
END_METHOD

METHOD GET_PSF : POINTER TO L_TB2P_scSF_TM_MotionControl
END_METHOD

METHOD ADDOFFSET
VAR_INPUT
	ITFTECHMODULE : L_TS2P_ISyncPosBase;
	LRSETPOS : LREAL;
	LRSETVEL : LREAL;
	LRSETOFFSET : LREAL;
	LRSETOFFSETVEL : LREAL;
	ETRAVERSINGRANGE : L_MC1P.L_MC1P_TraversingRange;
	LRCYCLELENGTH : LREAL;
END_VAR
VAR_OUTPUT
	XERROR : BOOL;
	EERRORID : L_IE1P.L_IE1P_Error;
	LRSETPOSOUT : LREAL;
	LRSETVELOUT : LREAL;
END_VAR
END_METHOD

METHOD CLUTCH
VAR_INPUT
	ITFTECHMODULE : L_TS2P_ISyncPosBase;
	XENABLE : BOOL;
	XSYNCIN : BOOL;
	LRSETBASEVELOCITY : LREAL;
	ESYNCMODE : L_TB2P_SyncMode;
	EALLOWEDDIRECTION : L_TB2P_AllowedDirection;
	LRSYNCVEL : LREAL;
	LRSYNCACC : LREAL;
	LRSYNCDEC : LREAL;
	LRSYNCJERK : LREAL;
	LRSYNCINDIST : LREAL;
	LRSYNCOUTDIST : LREAL;
	LRSYNCOUTPOS : LREAL;
	XLOADCLUTCHOFFSET : BOOL;
	LRLOADCLUTCHOFFSET : LREAL;
	LRCYCLICMASTERPOS : LREAL;
	LRCYCLICMASTERVEL : LREAL;
	ETRAVERSINGRANGEMASTER : L_MC1P_TraversingRange;
	LRCYCLELENGTHMASTER : LREAL;
	LRCYCLICAXISPOS : LREAL;
	LRCYCLICAXISVEL : LREAL;
	LRCYCLICAXISACC : LREAL;
	ETRAVERSINGRANGEAXIS : L_MC1P_TraversingRange;
	LRCYCLELENGTHAXIS : LREAL;
END_VAR
VAR_OUTPUT
	XERROR : BOOL;
	EERRORID : L_IE1P.L_IE1P_Error;
	XBUSY : BOOL;
	XDONE : BOOL;
	XSYNCHRONISED : BOOL;
	XACCDECSYNC : BOOL;
	XINBASEVELOCITY : BOOL;
	LRSETPOSOUT : LREAL;
	LRSETVELOUT : LREAL;
	LRSETACCOUT : LREAL;
	LRCLUTCHOFFSETOUT : LREAL;
END_VAR
END_METHOD

METHOD GEARBOX
VAR_INPUT
	ITFTECHMODULE : L_TS2P_ISyncPosBase;
	XENABLE : BOOL;
	LRSETPOSX : LREAL;
	LRSETVELX : LREAL;
	DWNUMERATOR : DWORD;
	DWDENOMINATOR : DWORD;
	LRCYCLELENGTHX : LREAL;
	LRCYCLELENGTHY : LREAL;
	ETRAVERSINGRANGEX : L_MC1P.L_MC1P_TraversingRange;
	ETRAVERSINGRANGEY : L_MC1P.L_MC1P_TraversingRange;
	XLOADGEARBOXPOS : BOOL;
	LRLOADGEARBOXPOS : LREAL;
END_VAR
VAR_OUTPUT
	XERROR : BOOL;
	EERRORID : L_IE1P.L_IE1P_Error;
	LRSETPOSOUT : LREAL;
	LRSETVELOUT : LREAL;
END_VAR
END_METHOD

METHOD OFFSETANDTRIM
VAR_INPUT
	ITFTECHMODULE : L_TS2P_ISyncPosBase;
	XENABLE : BOOL;
	LRSETOFFSET : LREAL;
	XTRIMPOS : BOOL;
	XTRIMNEG : BOOL;
	LRSETTRIMDISTANCE : LREAL;
	ETRIMMODE : L_TS2P_TrimMode;
	XLOADOFFSET : BOOL;
	XRESETTRIMOFFSET : BOOL;
	LRSETVEL : LREAL;
	LRSETACC : LREAL;
	LRSETDEC : LREAL;
	LRSETJERK : LREAL;
	WACTDIRECTION : WORD;
	EALLOWEDDIRECTION : L_TB2P.L_TB2P_AllowedDirection;
	LRCYCMASTERPOS : LREAL;
	LRCYCMASTERVEL : LREAL;
	LRCYCMASTERACC : LREAL;
END_VAR
VAR_OUTPUT
	XERROR : BOOL;
	EERRORID : L_IE1P.L_IE1P_Error;
	XBUSY : BOOL;
	XDONE : BOOL;
	LRSETOFFSETOUTTOTAL : LREAL;
	LRSETOFFSETOUTTOTALVEL : LREAL;
	LRSETOFFSETOUT : LREAL;
	LRSETOFFSETOUTTRIM : LREAL;
END_VAR
END_METHOD

METHOD REQUESTINTERFACE : BOOL
VAR_INPUT
	ID : DINT;
	PITFUNKNOWN : POINTER TO L_UBUP.L_UBUP_IUnknown;
END_VAR
END_METHOD

METHOD CALLFUNCTION
VAR_INPUT
	UIINPUTDATAIDX : UINT;
	UIOUTPUTDATAIDX : UINT;
END_VAR
END_METHOD

METHOD COPYINPUTS : BOOL
VAR_INPUT
	IDX : WORD;
END_VAR
END_METHOD

METHOD COPYOUTPUTS : BOOL
VAR_INPUT
	IDX : WORD;
END_VAR
END_METHOD

METHOD FUNCTIONWASCALLEDTWICE : BOOL
VAR_INPUT
	IDX : WORD;
END_VAR
END_METHOD

METHOD HANDLESTANDARDCALL : BOOL
END_METHOD

METHOD SYNCOUTPUTS
VAR_INPUT
	UICOPYOUTPUTFROMIDX : UINT;
	UICOPYOUTPUTTOIDX : UINT;
END_VAR
END_METHOD

METHOD FB_INIT : BOOL
VAR_INPUT
	BINITRETAINS : BOOL;
	BINCOPYCODE : BOOL;
END_VAR
END_METHOD

METHOD CALL_INTERNALCTRL
END_METHOD

(* ---- L_TS2P_SYNCRONISEDOVERRIDE.pou ---- *)
FUNCTION_BLOCK L_TS2P_SYNCRONISEDOVERRIDE
VAR_INPUT
	XENABLE : BOOL;
	XSYNCHRONISED : BOOL;
	XEXECUTEGAP : BOOL;
	XAUXEXECUTEGAP : BOOL;
	LRSYNCOVERRIDE : LREAL := 1;
	LRCYCMASTERPOS : LREAL;
	LRCYCMASTERVEL : LREAL;
	LRCYCMASTERACC : LREAL;
	LRCYCSLAVEPOS : LREAL;
	LRCYCSLAVEVEL : LREAL;
	LRCYCSLAVEACC : LREAL;
	LRACC : LREAL;
	LRDEC : LREAL;
	LRJERK : LREAL;
	LRTASKCYLCETIME : LREAL := 0.001;
END_VAR
VAR_OUTPUT
	XBUSY : BOOL;
	XERROR : BOOL;
	EERRORID : L_IE1P_Error;
	XOVERRIDELIMITED : BOOL;
	XEXECUTEGAPOUT : BOOL;
	XAUXEXECUTEGAPOUT : BOOL;
	LRSETPOS : LREAL;
	LRSETVEL : LREAL;
	LRSETACC : LREAL;
	XSYNCOVERRIDEACTIVE : BOOL;
	XRAMPGENBUSY : BOOL;
END_VAR
VAR
	XENABLE_OLD : BOOL;
	XEXECUTEGAP_OLD : BOOL;
	XAUXEXECUTEGAP_OLD : BOOL;
	LRSYNCOVERRIDE_INT : LREAL := 1;
	LRSYNCOVERRIDE_LOCK : LREAL;
	LRADDOVERRIDE_LOCK : LREAL;
	WSTATE : WORD := 0;
	LROFFSETPOS_INT : LREAL;
	LROFFSETVEL_INT : LREAL;
	LROFFSETACC_INT : LREAL;
	LROFFSETVEL_OLD : LREAL;
	LRVELTARGET : LREAL;
	LRVELSTART : LREAL;
	FB_RAMPGENERATOR1 : L_MC1P_RampGenerator;
	C_LRCYCLELENGTHMASTER : LREAL := (16#4FFFFFFFFFFFFFFF * 1E-08);
END_VAR
END_FUNCTION_BLOCK

METHOD CALL_ERRORHANDLER
END_METHOD

METHOD CALL_FB_RAMPGENERATOR1
END_METHOD

METHOD CALL_OUTPUTS
END_METHOD

METHOD CALL_RESETCOMMANDS
END_METHOD

METHOD CALL_RESETOUTPUTS
END_METHOD

METHOD CALL_STATEMACHINE
END_METHOD
